ABB RAPID module: Module1.mod

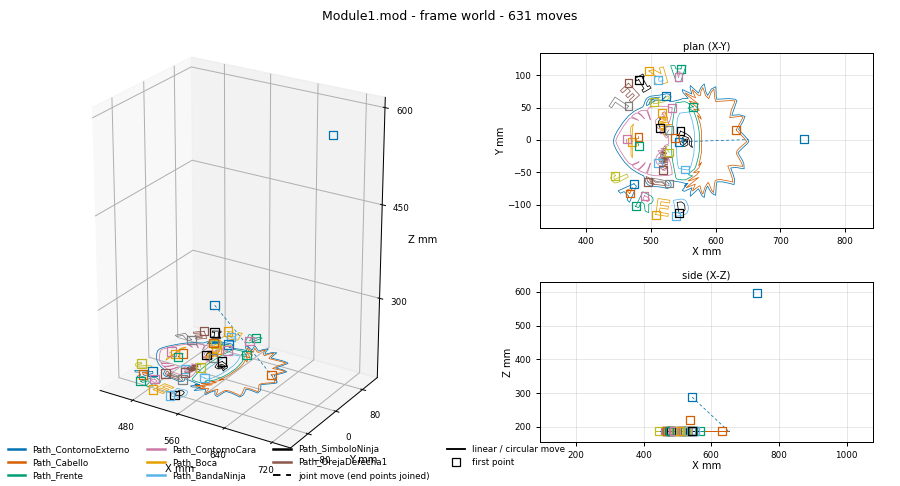
[picture p0: tool path of Module1.mod in frame world, 631 of 636 moves have a stored position in this frame; points joined in program order, loops and branches not executed]
MODULE Module1
    TASK PERS wobjdata Workobject_1:=[FALSE,TRUE,"",[[472.139180242,2.803580658,186.5],[0,0.573617827,0.819123061,0]],[[0,0,0],[1,0,0,0]]];
    TASK PERS wobjdata Cara:=[FALSE,TRUE,"",[[540.229,0.016,186.5],[0,0.707106781,0.707106781,0]],[[0,0,0],[1,0,0,0]]];
    PERS tooldata MyNewTool:=[TRUE,[[8.526,1.82,195.145],[0.965925826,0,0.258819045,0]],[0.14,[0,0,1],[1,0,0,0],0,0,0]];
    CONST robtarget Target_10:=[[-45.629166667,12.05,-2],[0.71519384,0,0,-0.698926156],[0,0,0,0],[9E+09,9E+09,9E+09,9E+09,9E+09,9E+09]];
    CONST robtarget Target_20:=[[-46.396458333,17.381354167,-2],[0.71519384,0,0,-0.698926156],[0,0,0,0],[9E+09,9E+09,9E+09,9E+09,9E+09,9E+09]];
    CONST robtarget Target_30:=[[-42.49468099,20.715104167,-2],[0.71519384,0,0,-0.698926156],[0,0,0,0],[9E+09,9E+09,9E+09,9E+09,9E+09,9E+09]];
    CONST robtarget Target_40:=[[-36.679635417,22.68625,-2],[0.71519384,0,0,-0.698926156],[0,0,0,0],[9E+09,9E+09,9E+09,9E+09,9E+09,9E+09]];
    CONST robtarget Target_50:=[[-21.710833333,26.072916667,-2],[0.71519384,0,0,-0.698926156],[0,0,0,0],[9E+09,9E+09,9E+09,9E+09,9E+09,9E+09]];
    CONST robtarget Target_60:=[[-4.75765625,27.104791667,-2],[0.71519384,0,0,-0.698926156],[0,0,0,0],[9E+09,9E+09,9E+09,9E+09,9E+09,9E+09]];
    CONST robtarget Target_70:=[[12.314583333,26.866666667,-2],[0.71519384,0,0,-0.698926156],[0,0,0,0],[9E+09,9E+09,9E+09,9E+09,9E+09,9E+09]];
    CONST robtarget Target_80:=[[26.688072917,24.458958333,-2],[0.71519384,0,0,-0.698926156],[0,0,0,0],[9E+09,9E+09,9E+09,9E+09,9E+09,9E+09]];
    CONST robtarget Target_90:=[[39.6725,20.46375,-2],[0.71519384,0,0,-0.698926156],[0,0,0,0],[9E+09,9E+09,9E+09,9E+09,9E+09,9E+09]];
    CONST robtarget Target_100:=[[43.257604167,18.849791667,-2],[0.71519384,0,0,-0.698926156],[0,0,0,0],[9E+09,9E+09,9E+09,9E+09,9E+09,9E+09]];
    CONST robtarget Target_110:=[[41.365833333,4.27125,-2],[0.71519384,0,0,-0.698926156],[0,0,0,0],[9E+09,9E+09,9E+09,9E+09,9E+09,9E+09]];
    CONST robtarget Target_120:=[[32.581666667,0.567083333,-2],[0.71519384,0,0,-0.698926156],[0,0,0,0],[9E+09,9E+09,9E+09,9E+09,9E+09,9E+09]];
    CONST robtarget Target_130:=[[22.252167969,-0.135716146,-2],[0.71519384,0,0,-0.698926156],[0,0,0,0],[9E+09,9E+09,9E+09,9E+09,9E+09,9E+09]];
    CONST robtarget Target_140:=[[-12.892766927,-0.549127604,-2],[0.71519384,0,0,-0.698926156],[0,0,0,0],[9E+09,9E+09,9E+09,9E+09,9E+09,9E+09]];
    CONST robtarget Target_150:=[[-26.05,-0.120833333,-2],[0.71519384,0,0,-0.698926156],[0,0,0,0],[9E+09,9E+09,9E+09,9E+09,9E+09,9E+09]];
    CONST robtarget Target_160:=[[-37.334479167,1.129322917,-2],[0.71519384,0,0,-0.698926156],[0,0,0,0],[9E+09,9E+09,9E+09,9E+09,9E+09,9E+09]];
    CONST robtarget Target_170:=[[-43.618333333,2.577916667,-2],[0.71519384,0,0,-0.698926156],[0,0,0,0],[9E+09,9E+09,9E+09,9E+09,9E+09,9E+09]];
    CONST robtarget Target_180:=[[-45.629166667,12.05,-2],[0.71519384,0,0,-0.698926156],[0,0,0,0],[9E+09,9E+09,9E+09,9E+09,9E+09,9E+09]];
    CONST robtarget Target_190:=[[0.514166667,109.68125,-2],[0.71519384,0,0,-0.698926156],[0,0,0,0],[9E+09,9E+09,9E+09,9E+09,9E+09,9E+09]];
    CONST robtarget Target_200:=[[16.547916667,95.129166667,-2],[0.71519384,0,0,-0.698926156],[0,0,0,0],[9E+09,9E+09,9E+09,9E+09,9E+09,9E+09]];
    CONST robtarget Target_210:=[[29.843229167,102.623489583,-2],[0.71519384,0,0,-0.698926156],[0,0,0,0],[9E+09,9E+09,9E+09,9E+09,9E+09,9E+09]];
    CONST robtarget Target_220:=[[36.33875,105.024583333,-2],[0.71519384,0,0,-0.698926156],[0,0,0,0],[9E+09,9E+09,9E+09,9E+09,9E+09,9E+09]];
    CONST robtarget Target_230:=[[38.865520833,96.729895833,-2],[0.71519384,0,0,-0.698926156],[0,0,0,0],[9E+09,9E+09,9E+09,9E+09,9E+09,9E+09]];
    CONST robtarget Target_240:=[[38.06515625,84.664895833,-2],[0.71519384,0,0,-0.698926156],[0,0,0,0],[9E+09,9E+09,9E+09,9E+09,9E+09,9E+09]];
    CONST robtarget Target_250:=[[60.680416667,92.642083333,-2],[0.71519384,0,0,-0.698926156],[0,0,0,0],[9E+09,9E+09,9E+09,9E+09,9E+09,9E+09]];
    CONST robtarget Target_260:=[[62.955833333,89.308333333,-2],[0.71519384,0,0,-0.698926156],[0,0,0,0],[9E+09,9E+09,9E+09,9E+09,9E+09,9E+09]];
    CONST robtarget Target_270:=[[63.82234375,79.750260417,-2],[0.71519384,0,0,-0.698926156],[0,0,0,0],[9E+09,9E+09,9E+09,9E+09,9E+09,9E+09]];
    CONST robtarget Target_280:=[[62.797083333,61.632916667,-2],[0.71519384,0,0,-0.698926156],[0,0,0,0],[9E+09,9E+09,9E+09,9E+09,9E+09,9E+09]];
    CONST robtarget Target_290:=[[67.427291667,60.640729167,-2],[0.71519384,0,0,-0.698926156],[0,0,0,0],[9E+09,9E+09,9E+09,9E+09,9E+09,9E+09]];
    CONST robtarget Target_300:=[[82.15796875,60.058645833,-2],[0.71519384,0,0,-0.698926156],[0,0,0,0],[9E+09,9E+09,9E+09,9E+09,9E+09,9E+09]];
    CONST robtarget Target_310:=[[78.797760417,53.338229167,-2],[0.71519384,0,0,-0.698926156],[0,0,0,0],[9E+09,9E+09,9E+09,9E+09,9E+09,9E+09]];
    CONST robtarget Target_320:=[[68.670833333,47.398333333,-2],[0.71519384,0,0,-0.698926156],[0,0,0,0],[9E+09,9E+09,9E+09,9E+09,9E+09,9E+09]];
    CONST robtarget Target_330:=[[74.352760417,44.5540625,-2],[0.71519384,0,0,-0.698926156],[0,0,0,0],[9E+09,9E+09,9E+09,9E+09,9E+09,9E+09]];
    CONST robtarget Target_340:=[[86.345,42.318333333,-2],[0.71519384,0,0,-0.698926156],[0,0,0,0],[9E+09,9E+09,9E+09,9E+09,9E+09,9E+09]];
    CONST robtarget Target_350:=[[84.1621875,39.53359375,-2],[0.71519384,0,0,-0.698926156],[0,0,0,0],[9E+09,9E+09,9E+09,9E+09,9E+09,9E+09]];
    CONST robtarget Target_360:=[[79.51875,36.232916667,-2],[0.71519384,0,0,-0.698926156],[0,0,0,0],[9E+09,9E+09,9E+09,9E+09,9E+09,9E+09]];
    CONST robtarget Target_370:=[[72.375,33.3225,-2],[0.71519384,0,0,-0.698926156],[0,0,0,0],[9E+09,9E+09,9E+09,9E+09,9E+09,9E+09]];
    CONST robtarget Target_380:=[[84.016666667,20.569583333,-2],[0.71519384,0,0,-0.698926156],[0,0,0,0],[9E+09,9E+09,9E+09,9E+09,9E+09,9E+09]];
    CONST robtarget Target_390:=[[80.821822917,20.331458333,-2],[0.71519384,0,0,-0.698926156],[0,0,0,0],[9E+09,9E+09,9E+09,9E+09,9E+09,9E+09]];
    CONST robtarget Target_400:=[[70.94625,22.950833333,-2],[0.71519384,0,0,-0.698926156],[0,0,0,0],[9E+09,9E+09,9E+09,9E+09,9E+09,9E+09]];
    CONST robtarget Target_410:=[[77.746041667,8.385520833,-2],[0.71519384,0,0,-0.698926156],[0,0,0,0],[9E+09,9E+09,9E+09,9E+09,9E+09,9E+09]];
    CONST robtarget Target_420:=[[73.598697917,9.146197917,-2],[0.71519384,0,0,-0.698926156],[0,0,0,0],[9E+09,9E+09,9E+09,9E+09,9E+09,9E+09]];
    CONST robtarget Target_430:=[[64.172916667,17.394583333,-2],[0.71519384,0,0,-0.698926156],[0,0,0,0],[9E+09,9E+09,9E+09,9E+09,9E+09,9E+09]];
    CONST robtarget Target_440:=[[63.736354167,8.65671875,-2],[0.71519384,0,0,-0.698926156],[0,0,0,0],[9E+09,9E+09,9E+09,9E+09,9E+09,9E+09]];
    CONST robtarget Target_450:=[[62.000852865,4.113326823,-2],[0.71519384,0,0,-0.698926156],[0,0,0,0],[9E+09,9E+09,9E+09,9E+09,9E+09,9E+09]];
    CONST robtarget Target_460:=[[59.28391276,-7.539915365,-2],[0.71519384,0,0,-0.698926156],[0,0,0,0],[9E+09,9E+09,9E+09,9E+09,9E+09,9E+09]];
    CONST robtarget Target_470:=[[58.987083333,-11.074583333,-2],[0.71519384,0,0,-0.698926156],[0,0,0,0],[9E+09,9E+09,9E+09,9E+09,9E+09,9E+09]];
    CONST robtarget Target_480:=[[66.7790625,-9.156354167,-2],[0.71519384,0,0,-0.698926156],[0,0,0,0],[9E+09,9E+09,9E+09,9E+09,9E+09,9E+09]];
    CONST robtarget Target_490:=[[70.522916667,-12.027083333,-2],[0.715023643,0.015246994,0.015601871,-0.69875983],[0,0,0,0],[9E+09,9E+09,9E+09,9E+09,9E+09,9E+09]];
    CONST robtarget Target_500:=[[71.26375,-15.744479167,-2],[0.714513134,0.030486731,0.031196317,-0.698260933],[0,0,0,0],[9E+09,9E+09,9E+09,9E+09,9E+09,9E+09]];
    CONST robtarget Target_510:=[[69.391822917,-25.586979167,-2],[0.713662555,0.045711958,0.046775915,-0.697429701],[0,0,0,0],[9E+09,9E+09,9E+09,9E+09,9E+09,9E+09]];
    CONST robtarget Target_520:=[[67.380989583,-41.475208333,-2],[0.712472311,0.060915428,0.06233325,-0.696266531],[0,0,0,0],[9E+09,9E+09,9E+09,9E+09,9E+09,9E+09]];
    CONST robtarget Target_530:=[[64.490416667,-46.158333333,-2],[0.712472311,0.060915428,0.06233325,-0.696266531],[0,0,0,0],[9E+09,9E+09,9E+09,9E+09,9E+09,9E+09]];
    CONST robtarget Target_540:=[[61.67921875,-48.387447917,-2],[0.712472311,0.060915428,0.06233325,-0.696266531],[0,0,0,0],[9E+09,9E+09,9E+09,9E+09,9E+09,9E+09]];
    CONST robtarget Target_550:=[[54.350260417,-51.03328125,-2],[0.712472311,0.060915428,0.06233325,-0.696266531],[0,0,0,0],[9E+09,9E+09,9E+09,9E+09,9E+09,9E+09]];
    CONST robtarget Target_560:=[[51.214947917,-52.409114583,-2],[0.710942969,0.076089906,0.077860918,-0.694771976],[0,0,0,0],[9E+09,9E+09,9E+09,9E+09,9E+09,9E+09]];
    CONST robtarget Target_570:=[[44.472207031,-65.71186849,-2],[0.710942969,0.076089906,0.077860918,-0.694771976],[0,0,0,0],[9E+09,9E+09,9E+09,9E+09,9E+09,9E+09]];
    CONST robtarget Target_580:=[[37.364010417,-74.52828125,-2],[0.710942969,0.076089906,0.077860918,-0.694771976],[0,0,0,0],[9E+09,9E+09,9E+09,9E+09,9E+09,9E+09]];
    CONST robtarget Target_590:=[[27.586829427,-82.957740885,-2],[0.706870064,0.106323014,0.108797708,-0.690791712],[0,0,0,0],[9E+09,9E+09,9E+09,9E+09,9E+09,9E+09]];
    CONST robtarget Target_600:=[[14.43125,-91.719583333,-2],[0.709075257,0.09122817,0.093351528,-0.692946746],[0,0,0,0],[9E+09,9E+09,9E+09,9E+09,9E+09,9E+09]];
    CONST robtarget Target_610:=[[5.091458333,-96.535,-2],[0.709075257,0.09122817,0.093351528,-0.692946746],[0,0,0,0],[9E+09,9E+09,9E+09,9E+09,9E+09,9E+09]];
    CONST robtarget Target_620:=[[-1.867083333,-98.016666667,-2],[0.709075257,0.09122817,0.093351528,-0.692946746],[0,0,0,0],[9E+09,9E+09,9E+09,9E+09,9E+09,9E+09]];
    CONST robtarget Target_630:=[[-7.6746875,-97.037708333,-2],[0.709075257,0.09122817,0.093351528,-0.692946746],[0,0,0,0],[9E+09,9E+09,9E+09,9E+09,9E+09,9E+09]];
    CONST robtarget Target_640:=[[-16.101666667,-93.095416667,-2],[0.709075257,0.09122817,0.093351528,-0.692946746],[0,0,0,0],[9E+09,9E+09,9E+09,9E+09,9E+09,9E+09]];
    CONST robtarget Target_650:=[[-24.727083333,-87.6846875,-2],[0.709075257,0.09122817,0.093351528,-0.692946746],[0,0,0,0],[9E+09,9E+09,9E+09,9E+09,9E+09,9E+09]];
    CONST robtarget Target_660:=[[-35.09875,-80.130833333,-2],[0.710942969,0.076089907,0.077860918,-0.694771976],[0,0,0,0],[9E+09,9E+09,9E+09,9E+09,9E+09,9E+09]];
    CONST robtarget Target_670:=[[-44.36578125,-70.652135417,-2],[0.712472311,0.060915428,0.06233325,-0.696266531],[0,0,0,0],[9E+09,9E+09,9E+09,9E+09,9E+09,9E+09]];
    CONST robtarget Target_680:=[[-50.97375,-60.34,-2],[0.712472311,0.060915428,0.06233325,-0.696266531],[0,0,0,0],[9E+09,9E+09,9E+09,9E+09,9E+09,9E+09]];
    CONST robtarget Target_690:=[[-55.41875,-51.29125,-2],[0.712989136,0.054837114,0.056113461,-0.6967716],[0,0,0,0],[9E+09,9E+09,9E+09,9E+09,9E+09,9E+09]];
    CONST robtarget Target_700:=[[-66.055,-47.434947917,-2],[0.712989136,0.054837114,0.05611346,-0.6967716],[0,0,0,0],[9E+09,9E+09,9E+09,9E+09,9E+09,9E+09]];
    CONST robtarget Target_710:=[[-69.124166667,-44.570833333,-2],[0.713662554,0.045711958,0.046775915,-0.697429702],[0,0,0,0],[9E+09,9E+09,9E+09,9E+09,9E+09,9E+09]];
    CONST robtarget Target_720:=[[-71.03578125,-40.092760417,-2],[0.714513134,0.030486731,0.031196317,-0.698260933],[0,0,0,0],[9E+09,9E+09,9E+09,9E+09,9E+09,9E+09]];
    CONST robtarget Target_730:=[[-72.735729167,-24.707239583,-2],[0.71519384,0,0,-0.698926156],[0,0,0,0],[9E+09,9E+09,9E+09,9E+09,9E+09,9E+09]];
    CONST robtarget Target_740:=[[-74.733333333,-14.9375,-2],[0.71519384,0,0,-0.698926156],[0,0,0,0],[9E+09,9E+09,9E+09,9E+09,9E+09,9E+09]];
    CONST robtarget Target_750:=[[-73.57578125,-11.312708333,-2],[0.71519384,0,0,-0.698926156],[0,0,0,0],[9E+09,9E+09,9E+09,9E+09,9E+09,9E+09]];
    CONST robtarget Target_760:=[[-71.029166667,-8.957916667,-2],[0.71519384,0,0,-0.698926156],[0,0,0,0],[9E+09,9E+09,9E+09,9E+09,9E+09,9E+09]];
    CONST robtarget Target_770:=[[-67.4440625,-9.1034375,-2],[0.71519384,0,0,-0.698926156],[0,0,0,0],[9E+09,9E+09,9E+09,9E+09,9E+09,9E+09]];
    CONST robtarget Target_780:=[[-63.03875,-11.7625,-2],[0.71519384,0,0,-0.698926156],[0,0,0,0],[9E+09,9E+09,9E+09,9E+09,9E+09,9E+09]];
    CONST robtarget Target_790:=[[-62.873385417,-8.045104167,-2],[0.71519384,0,0,-0.698926156],[0,0,0,0],[9E+09,9E+09,9E+09,9E+09,9E+09,9E+09]];
    CONST robtarget Target_800:=[[-65.347239583,7.22796875,-2],[0.71519384,0,0,-0.698926156],[0,0,0,0],[9E+09,9E+09,9E+09,9E+09,9E+09,9E+09]];
    CONST robtarget Target_810:=[[-66.795833333,11.838333333,-2],[0.71519384,0,0,-0.698926156],[0,0,0,0],[9E+09,9E+09,9E+09,9E+09,9E+09,9E+09]];
    CONST robtarget Target_820:=[[-67.272083333,15.225,-2],[0.71519384,0,0,-0.698926156],[0,0,0,0],[9E+09,9E+09,9E+09,9E+09,9E+09,9E+09]];
    CONST robtarget Target_830:=[[-71.29375,11.785416667,-2],[0.71519384,0,0,-0.698926156],[0,0,0,0],[9E+09,9E+09,9E+09,9E+09,9E+09,9E+09]];
    CONST robtarget Target_840:=[[-66.4915625,17.024166667,-2],[0.71519384,0,0,-0.698926156],[0,0,0,0],[9E+09,9E+09,9E+09,9E+09,9E+09,9E+09]];
    CONST robtarget Target_850:=[[-77.769427083,8.286302083,-2],[0.71519384,0,0,-0.698926156],[0,0,0,0],[9E+09,9E+09,9E+09,9E+09,9E+09,9E+09]];
    CONST robtarget Target_860:=[[-79.264322917,11.408385417,-2],[0.71519384,0,0,-0.698926156],[0,0,0,0],[9E+09,9E+09,9E+09,9E+09,9E+09,9E+09]];
    CONST robtarget Target_870:=[[-73.780833333,23.1625,-2],[0.71519384,0,0,-0.698926156],[0,0,0,0],[9E+09,9E+09,9E+09,9E+09,9E+09,9E+09]];
    CONST robtarget Target_880:=[[-81.923385417,20.609270833,-2],[0.71519384,0,0,-0.698926156],[0,0,0,0],[9E+09,9E+09,9E+09,9E+09,9E+09,9E+09]];
    CONST robtarget Target_890:=[[-86.904166667,20.6225,-2],[0.71519384,0,0,-0.698926156],[0,0,0,0],[9E+09,9E+09,9E+09,9E+09,9E+09,9E+09]];
    CONST robtarget Target_900:=[[-75.2625,33.269583333,-2],[0.71519384,0,0,-0.698926156],[0,0,0,0],[9E+09,9E+09,9E+09,9E+09,9E+09,9E+09]];
    CONST robtarget Target_910:=[[-86.203020833,38.7596875,-2],[0.71519384,0,0,-0.698926156],[0,0,0,0],[9E+09,9E+09,9E+09,9E+09,9E+09,9E+09]];
    CONST robtarget Target_920:=[[-88.809166667,42.159583333,-2],[0.71519384,0,0,-0.698926156],[0,0,0,0],[9E+09,9E+09,9E+09,9E+09,9E+09,9E+09]];
    CONST robtarget Target_930:=[[-80.170520833,43.555260417,-2],[0.71519384,0,0,-0.698926156],[0,0,0,0],[9E+09,9E+09,9E+09,9E+09,9E+09,9E+09]];
    CONST robtarget Target_940:=[[-73.9925,45.599166667,-2],[0.71519384,0,0,-0.698926156],[0,0,0,0],[9E+09,9E+09,9E+09,9E+09,9E+09,9E+09]];
    CONST robtarget Target_950:=[[-71.23421875,47.2528125,-2],[0.71519384,0,0,-0.698926156],[0,0,0,0],[9E+09,9E+09,9E+09,9E+09,9E+09,9E+09]];
    CONST robtarget Target_960:=[[-76.479583333,50.077239583,-2],[0.71519384,0,0,-0.698926156],[0,0,0,0],[9E+09,9E+09,9E+09,9E+09,9E+09,9E+09]];
    CONST robtarget Target_970:=[[-81.506666667,53.272083333,-2],[0.71519384,0,0,-0.698926156],[0,0,0,0],[9E+09,9E+09,9E+09,9E+09,9E+09,9E+09]];
    CONST robtarget Target_980:=[[-84.026822917,56.665364583,-2],[0.71519384,0,0,-0.698926156],[0,0,0,0],[9E+09,9E+09,9E+09,9E+09,9E+09,9E+09]];
    CONST robtarget Target_990:=[[-85.316666667,59.622083333,-2],[0.71519384,0,0,-0.698926156],[0,0,0,0],[9E+09,9E+09,9E+09,9E+09,9E+09,9E+09]];
    CONST robtarget Target_1000:=[[-78.860833333,60.15125,-2],[0.71519384,0,0,-0.698926156],[0,0,0,0],[9E+09,9E+09,9E+09,9E+09,9E+09,9E+09]];
    CONST robtarget Target_1010:=[[-69.501197917,60.706875,-2],[0.71519384,0,0,-0.698926156],[0,0,0,0],[9E+09,9E+09,9E+09,9E+09,9E+09,9E+09]];
    CONST robtarget Target_1020:=[[-64.62625,61.8975,-2],[0.71519384,0,0,-0.698926156],[0,0,0,0],[9E+09,9E+09,9E+09,9E+09,9E+09,9E+09]];
    CONST robtarget Target_1030:=[[-64.619635417,70.126041667,-2],[0.71519384,0,0,-0.698926156],[0,0,0,0],[9E+09,9E+09,9E+09,9E+09,9E+09,9E+09]];
    CONST robtarget Target_1040:=[[-67.272083333,82.323333333,-2],[0.71519384,0,0,-0.698926156],[0,0,0,0],[9E+09,9E+09,9E+09,9E+09,9E+09,9E+09]];
    CONST robtarget Target_1050:=[[-68.9125,87.985416667,-2],[0.71519384,0,0,-0.698926156],[0,0,0,0],[9E+09,9E+09,9E+09,9E+09,9E+09,9E+09]];
    CONST robtarget Target_1060:=[[-62.297916667,89.149583333,-2],[0.71519384,0,0,-0.698926156],[0,0,0,0],[9E+09,9E+09,9E+09,9E+09,9E+09,9E+09]];
    CONST robtarget Target_1070:=[[-54.677916667,87.2975,-2],[0.71519384,0,0,-0.698926156],[0,0,0,0],[9E+09,9E+09,9E+09,9E+09,9E+09,9E+09]];
    CONST robtarget Target_1080:=[[-43.280989583,82.95171875,-2],[0.71519384,0,0,-0.698926156],[0,0,0,0],[9E+09,9E+09,9E+09,9E+09,9E+09,9E+09]];
    CONST robtarget Target_1090:=[[-42.275572917,90.479114583,-2],[0.71519384,0,0,-0.698926156],[0,0,0,0],[9E+09,9E+09,9E+09,9E+09,9E+09,9E+09]];
    CONST robtarget Target_1100:=[[-44.570833333,103.754583333,-2],[0.71519384,0,0,-0.698926156],[0,0,0,0],[9E+09,9E+09,9E+09,9E+09,9E+09,9E+09]];
    CONST robtarget Target_1110:=[[-36.633333333,103.278333333,-2],[0.71519384,0,0,-0.698926156],[0,0,0,0],[9E+09,9E+09,9E+09,9E+09,9E+09,9E+09]];
    CONST robtarget Target_1120:=[[-31.381354167,101.055833333,-2],[0.71519384,0,0,-0.698926156],[0,0,0,0],[9E+09,9E+09,9E+09,9E+09,9E+09,9E+09]];
    CONST robtarget Target_1130:=[[-19.752916667,94.070833333,-2],[0.71519384,0,0,-0.698926156],[0,0,0,0],[9E+09,9E+09,9E+09,9E+09,9E+09,9E+09]];
    CONST robtarget Target_1140:=[[-13.918854167,99.69984375,-2],[0.71519384,0,0,-0.698926156],[0,0,0,0],[9E+09,9E+09,9E+09,9E+09,9E+09,9E+09]];
    CONST robtarget Target_1150:=[[-6.259166667,107.987916667,-2],[0.71519384,0,0,-0.698926156],[0,0,0,0],[9E+09,9E+09,9E+09,9E+09,9E+09,9E+09]];
    CONST robtarget Target_1160:=[[-2.93203125,110.858645833,-2],[0.71519384,0,0,-0.698926156],[0,0,0,0],[9E+09,9E+09,9E+09,9E+09,9E+09,9E+09]];
    CONST robtarget Target_1170:=[[0.514166667,109.68125,-2],[0.71519384,0,0,-0.698926156],[0,0,0,0],[9E+09,9E+09,9E+09,9E+09,9E+09,9E+09]];
    CONST robtarget Target_1350:=[[15.489583333,91.425,-2],[0.71519384,0,0,-0.698926156],[0,0,0,0],[9E+09,9E+09,9E+09,9E+09,9E+09,9E+09]];
    CONST robtarget Target_1360:=[[34.94389974,101.979394531,-2],[0.71519384,0,0,-0.698926156],[0,0,0,0],[9E+09,9E+09,9E+09,9E+09,9E+09,9E+09]];
    CONST robtarget Target_1370:=[[36.669479167,98.674583333,-2],[0.71519384,0,0,-0.698926156],[0,0,0,0],[9E+09,9E+09,9E+09,9E+09,9E+09,9E+09]];
    CONST robtarget Target_1380:=[[34.321302083,81.436979167,-2],[0.71519384,0,0,-0.698926156],[0,0,0,0],[9E+09,9E+09,9E+09,9E+09,9E+09,9E+09]];
    CONST robtarget Target_1390:=[[46.763333333,84.016666667,-2],[0.71519384,0,0,-0.698926156],[0,0,0,0],[9E+09,9E+09,9E+09,9E+09,9E+09,9E+09]];
    CONST robtarget Target_1400:=[[56.129583333,88.177239583,-2],[0.71519384,0,0,-0.698926156],[0,0,0,0],[9E+09,9E+09,9E+09,9E+09,9E+09,9E+09]];
    CONST robtarget Target_1410:=[[60.257083333,89.52,-2],[0.71519384,0,0,-0.698926156],[0,0,0,0],[9E+09,9E+09,9E+09,9E+09,9E+09,9E+09]];
    CONST robtarget Target_1420:=[[60.706875,81.291458333,-2],[0.71519384,0,0,-0.698926156],[0,0,0,0],[9E+09,9E+09,9E+09,9E+09,9E+09,9E+09]];
    CONST robtarget Target_1430:=[[59.304583333,59.886666667,-2],[0.71519384,0,0,-0.698926156],[0,0,0,0],[9E+09,9E+09,9E+09,9E+09,9E+09,9E+09]];
    CONST robtarget Target_1440:=[[63.8025,58.56375,-2],[0.71519384,0,0,-0.698926156],[0,0,0,0],[9E+09,9E+09,9E+09,9E+09,9E+09,9E+09]];
    CONST robtarget Target_1450:=[[78.725,57.029166667,-2],[0.71519384,0,0,-0.698926156],[0,0,0,0],[9E+09,9E+09,9E+09,9E+09,9E+09,9E+09]];
    CONST robtarget Target_1460:=[[73.48625,52.84875,-2],[0.71519384,0,0,-0.698926156],[0,0,0,0],[9E+09,9E+09,9E+09,9E+09,9E+09,9E+09]];
    CONST robtarget Target_1470:=[[63.709895833,49.151197917,-2],[0.71519384,0,0,-0.698926156],[0,0,0,0],[9E+09,9E+09,9E+09,9E+09,9E+09,9E+09]];
    CONST robtarget Target_1480:=[[68.50546875,44.21671875,-2],[0.71519384,0,0,-0.698926156],[0,0,0,0],[9E+09,9E+09,9E+09,9E+09,9E+09,9E+09]];
    CONST robtarget Target_1490:=[[80.861510417,40.042916667,-2],[0.71519384,0,0,-0.698926156],[0,0,0,0],[9E+09,9E+09,9E+09,9E+09,9E+09,9E+09]];
    CONST robtarget Target_1500:=[[75.655833333,37.238333333,-2],[0.71519384,0,0,-0.698926156],[0,0,0,0],[9E+09,9E+09,9E+09,9E+09,9E+09,9E+09]];
    CONST robtarget Target_1510:=[[68.466608073,36.107239583,-2],[0.71519384,0,0,-0.698926156],[0,0,0,0],[9E+09,9E+09,9E+09,9E+09,9E+09,9E+09]];
    CONST robtarget Target_1520:=[[69.142949219,32.819791667,-2],[0.71519384,0,0,-0.698926156],[0,0,0,0],[9E+09,9E+09,9E+09,9E+09,9E+09,9E+09]];
    CONST robtarget Target_1530:=[[77.507916667,23.850416667,-2],[0.71519384,0,0,-0.698926156],[0,0,0,0],[9E+09,9E+09,9E+09,9E+09,9E+09,9E+09]];
    CONST robtarget Target_1540:=[[74.504895833,24.544947917,-2],[0.71519384,0,0,-0.698926156],[0,0,0,0],[9E+09,9E+09,9E+09,9E+09,9E+09,9E+09]];
    CONST robtarget Target_1550:=[[65.0725,28.771666667,-2],[0.71519384,0,0,-0.698926156],[0,0,0,0],[9E+09,9E+09,9E+09,9E+09,9E+09,9E+09]];
    CONST robtarget Target_1560:=[[67.03703125,24.128229167,-2],[0.71519384,0,0,-0.698926156],[0,0,0,0],[9E+09,9E+09,9E+09,9E+09,9E+09,9E+09]];
    CONST robtarget Target_1570:=[[72.6925,12.685,-2],[0.71519384,0,0,-0.698926156],[0,0,0,0],[9E+09,9E+09,9E+09,9E+09,9E+09,9E+09]];
    CONST robtarget Target_1580:=[[69.028020833,15.992291667,-2],[0.71519384,0,0,-0.698926156],[0,0,0,0],[9E+09,9E+09,9E+09,9E+09,9E+09,9E+09]];
    CONST robtarget Target_1590:=[[55.124166667,33.587083333,-2],[0.71519384,0,0,-0.698926156],[0,0,0,0],[9E+09,9E+09,9E+09,9E+09,9E+09,9E+09]];
    CONST robtarget Target_1600:=[[60.376145833,19.008541667,-2],[0.71519384,0,0,-0.698926156],[0,0,0,0],[9E+09,9E+09,9E+09,9E+09,9E+09,9E+09]];
    CONST robtarget Target_1610:=[[57.267291667,21.660989583,-2],[0.71519384,0,0,-0.698926156],[0,0,0,0],[9E+09,9E+09,9E+09,9E+09,9E+09,9E+09]];
    CONST robtarget Target_1620:=[[53.272083333,27.554583333,-2],[0.71519384,0,0,-0.698926156],[0,0,0,0],[9E+09,9E+09,9E+09,9E+09,9E+09,9E+09]];
    CONST robtarget Target_1630:=[[48.787395833,32.297239583,-2],[0.71519384,0,0,-0.698926156],[0,0,0,0],[9E+09,9E+09,9E+09,9E+09,9E+09,9E+09]];
    CONST robtarget Target_1640:=[[45.652083333,34.698333333,-2],[0.71519384,0,0,-0.698926156],[0,0,0,0],[9E+09,9E+09,9E+09,9E+09,9E+09,9E+09]];
    CONST robtarget Target_1650:=[[47.656302083,25.771126302,-2],[0.71519384,0,0,-0.698926156],[0,0,0,0],[9E+09,9E+09,9E+09,9E+09,9E+09,9E+09]];
    CONST robtarget Target_1660:=[[41.471666667,32.581666667,-2],[0.71519384,0,0,-0.698926156],[0,0,0,0],[9E+09,9E+09,9E+09,9E+09,9E+09,9E+09]];
    CONST robtarget Target_1670:=[[36.18,36.193229167,-2],[0.71519384,0,0,-0.698926156],[0,0,0,0],[9E+09,9E+09,9E+09,9E+09,9E+09,9E+09]];
    CONST robtarget Target_1680:=[[31.957725423,37.723368327,-2],[0.71519384,0,0,-0.698926156],[0,0,0,0],[9E+09,9E+09,9E+09,9E+09,9E+09,9E+09]];
    CONST robtarget Target_1690:=[[38.137916667,31.787916667,-2],[0.71519384,0,0,-0.698926156],[0,0,0,0],[9E+09,9E+09,9E+09,9E+09,9E+09,9E+09]];
    CONST robtarget Target_1700:=[[24.262174479,36.184960938,-2],[0.71519384,0,0,-0.698926156],[0,0,0,0],[9E+09,9E+09,9E+09,9E+09,9E+09,9E+09]];
    CONST robtarget Target_1710:=[[11.282708333,38.2040625,-2],[0.71519384,0,0,-0.698926156],[0,0,0,0],[9E+09,9E+09,9E+09,9E+09,9E+09,9E+09]];
    CONST robtarget Target_1720:=[[-18.377083333,37.92625,-2],[0.71519384,0,0,-0.698926156],[0,0,0,0],[9E+09,9E+09,9E+09,9E+09,9E+09,9E+09]];
    CONST robtarget Target_1730:=[[-27.955,36.265989583,-2],[0.71519384,0,0,-0.698926156],[0,0,0,0],[9E+09,9E+09,9E+09,9E+09,9E+09,9E+09]];
    CONST robtarget Target_1740:=[[-39.328052572,33.621809896,-2],[0.71519384,0,0,-0.698926156],[0,0,0,0],[9E+09,9E+09,9E+09,9E+09,9E+09,9E+09]];
    CONST robtarget Target_1750:=[[-34.252083333,38.085,-2],[0.71519384,0,0,-0.698926156],[0,0,0,0],[9E+09,9E+09,9E+09,9E+09,9E+09,9E+09]];
    CONST robtarget Target_1760:=[[-42.851041667,34.01703125,-2],[0.71519384,0,0,-0.698926156],[0,0,0,0],[9E+09,9E+09,9E+09,9E+09,9E+09,9E+09]];
    CONST robtarget Target_1770:=[[-50.644054362,25.739603678,-2],[0.71519384,0,0,-0.698926156],[0,0,0,0],[9E+09,9E+09,9E+09,9E+09,9E+09,9E+09]];
    CONST robtarget Target_1780:=[[-48.539583333,34.698333333,-2],[0.71519384,0,0,-0.698926156],[0,0,0,0],[9E+09,9E+09,9E+09,9E+09,9E+09,9E+09]];
    CONST robtarget Target_1790:=[[-53.6725,30.729583333,-2],[0.71519384,0,0,-0.698926156],[0,0,0,0],[9E+09,9E+09,9E+09,9E+09,9E+09,9E+09]];
    CONST robtarget Target_1800:=[[-61.329707031,20.051165365,-2],[0.71519384,0,0,-0.698926156],[0,0,0,0],[9E+09,9E+09,9E+09,9E+09,9E+09,9E+09]];
    CONST robtarget Target_1810:=[[-62.9990625,17.354895833,-2],[0.71519384,0,0,-0.698926156],[0,0,0,0],[9E+09,9E+09,9E+09,9E+09,9E+09,9E+09]];
    CONST robtarget Target_1820:=[[-62.78078125,20.64234375,-2],[0.71519384,0,0,-0.698926156],[0,0,0,0],[9E+09,9E+09,9E+09,9E+09,9E+09,9E+09]];
    CONST robtarget Target_1830:=[[-57.890020345,33.671419271,-2],[0.71519384,0,0,-0.698926156],[0,0,0,0],[9E+09,9E+09,9E+09,9E+09,9E+09,9E+09]];
    CONST robtarget Target_1840:=[[-71.141614583,17.163072917,-2],[0.71519384,0,0,-0.698926156],[0,0,0,0],[9E+09,9E+09,9E+09,9E+09,9E+09,9E+09]];
    CONST robtarget Target_1850:=[[-73.87922526,14.268365885,-2],[0.71519384,0,0,-0.698926156],[0,0,0,0],[9E+09,9E+09,9E+09,9E+09,9E+09,9E+09]];
    CONST robtarget Target_1860:=[[-70.215572917,23.030208333,-2],[0.71519384,0,0,-0.698926156],[0,0,0,0],[9E+09,9E+09,9E+09,9E+09,9E+09,9E+09]];
    CONST robtarget Target_1870:=[[-68.184895833,28.407864583,-2],[0.71519384,0,0,-0.698926156],[0,0,0,0],[9E+09,9E+09,9E+09,9E+09,9E+09,9E+09]];
    CONST robtarget Target_1880:=[[-78.65578125,24.088541667,-2],[0.71519384,0,0,-0.698926156],[0,0,0,0],[9E+09,9E+09,9E+09,9E+09,9E+09,9E+09]];
    CONST robtarget Target_1890:=[[-72.080885417,32.7271875,-2],[0.71519384,0,0,-0.698926156],[0,0,0,0],[9E+09,9E+09,9E+09,9E+09,9E+09,9E+09]];
    CONST robtarget Target_1900:=[[-70.65875,35.650833333,-2],[0.71519384,0,0,-0.698926156],[0,0,0,0],[9E+09,9E+09,9E+09,9E+09,9E+09,9E+09]];
    CONST robtarget Target_1910:=[[-80.018385417,37.979166667,-2],[0.71519384,0,0,-0.698926156],[0,0,0,0],[9E+09,9E+09,9E+09,9E+09,9E+09,9E+09]];
    CONST robtarget Target_1920:=[[-83.570416667,39.884166667,-2],[0.71519384,0,0,-0.698926156],[0,0,0,0],[9E+09,9E+09,9E+09,9E+09,9E+09,9E+09]];
    CONST robtarget Target_1930:=[[-72.041197917,43.74046875,-2],[0.71519384,0,0,-0.698926156],[0,0,0,0],[9E+09,9E+09,9E+09,9E+09,9E+09,9E+09]];
    CONST robtarget Target_1940:=[[-65.26125,48.192083333,-2],[0.71519384,0,0,-0.698926156],[0,0,0,0],[9E+09,9E+09,9E+09,9E+09,9E+09,9E+09]];
    CONST robtarget Target_1950:=[[-68.965416667,50.15,-2],[0.71519384,0,0,-0.698926156],[0,0,0,0],[9E+09,9E+09,9E+09,9E+09,9E+09,9E+09]];
    CONST robtarget Target_1960:=[[-77.564375,53.589583333,-2],[0.71519384,0,0,-0.698926156],[0,0,0,0],[9E+09,9E+09,9E+09,9E+09,9E+09,9E+09]];
    CONST robtarget Target_1970:=[[-81.244150391,56.486150716,-2],[0.71519384,0,0,-0.698926156],[0,0,0,0],[9E+09,9E+09,9E+09,9E+09,9E+09,9E+09]];
    CONST robtarget Target_1980:=[[-67.42421875,58.02796875,-2],[0.71519384,0,0,-0.698926156],[0,0,0,0],[9E+09,9E+09,9E+09,9E+09,9E+09,9E+09]];
    CONST robtarget Target_1990:=[[-63.144583333,59.145833333,-2],[0.71519384,0,0,-0.698926156],[0,0,0,0],[9E+09,9E+09,9E+09,9E+09,9E+09,9E+09]];
    CONST robtarget Target_2000:=[[-61.466959635,61.796627604,-2],[0.71519384,0,0,-0.698926156],[0,0,0,0],[9E+09,9E+09,9E+09,9E+09,9E+09,9E+09]];
    CONST robtarget Target_2010:=[[-60.95515625,66.7790625,-2],[0.71519384,0,0,-0.698926156],[0,0,0,0],[9E+09,9E+09,9E+09,9E+09,9E+09,9E+09]];
    CONST robtarget Target_2020:=[[-63.409166667,80.206666667,-2],[0.71519384,0,0,-0.698926156],[0,0,0,0],[9E+09,9E+09,9E+09,9E+09,9E+09,9E+09]];
    CONST robtarget Target_2030:=[[-65.049583333,86.50375,-2],[0.71519384,0,0,-0.698926156],[0,0,0,0],[9E+09,9E+09,9E+09,9E+09,9E+09,9E+09]];
    CONST robtarget Target_2040:=[[-58.408541667,85.240364583,-2],[0.71519384,0,0,-0.698926156],[0,0,0,0],[9E+09,9E+09,9E+09,9E+09,9E+09,9E+09]];
    CONST robtarget Target_2050:=[[-47.9575,81.635416667,-2],[0.71519384,0,0,-0.698926156],[0,0,0,0],[9E+09,9E+09,9E+09,9E+09,9E+09,9E+09]];
    CONST robtarget Target_2060:=[[-40.258125,78.42734375,-2],[0.71519384,0,0,-0.698926156],[0,0,0,0],[9E+09,9E+09,9E+09,9E+09,9E+09,9E+09]];
    CONST robtarget Target_2070:=[[-38.80953125,85.743072917,-2],[0.71519384,0,0,-0.698926156],[0,0,0,0],[9E+09,9E+09,9E+09,9E+09,9E+09,9E+09]];
    CONST robtarget Target_2080:=[[-40.81375,101.796666667,-2],[0.71519384,0,0,-0.698926156],[0,0,0,0],[9E+09,9E+09,9E+09,9E+09,9E+09,9E+09]];
    CONST robtarget Target_2090:=[[-35.389791667,99.68,-2],[0.71519384,0,0,-0.698926156],[0,0,0,0],[9E+09,9E+09,9E+09,9E+09,9E+09,9E+09]];
    CONST robtarget Target_2100:=[[-21.492552083,91.92109375,-2],[0.71519384,0,0,-0.698926156],[0,0,0,0],[9E+09,9E+09,9E+09,9E+09,9E+09,9E+09]];
    CONST robtarget Target_2110:=[[-16.706074219,92.589166667,-2],[0.71519384,0,0,-0.698926156],[0,0,0,0],[9E+09,9E+09,9E+09,9E+09,9E+09,9E+09]];
    CONST robtarget Target_2120:=[[-12.787760417,96.121354167,-2],[0.71519384,0,0,-0.698926156],[0,0,0,0],[9E+09,9E+09,9E+09,9E+09,9E+09,9E+09]];
    CONST robtarget Target_2130:=[[-2.555,107.829166667,-2],[0.71519384,0,0,-0.698926156],[0,0,0,0],[9E+09,9E+09,9E+09,9E+09,9E+09,9E+09]];
    CONST robtarget Target_2140:=[[2.604375,103.90671875,-2],[0.71519384,0,0,-0.698926156],[0,0,0,0],[9E+09,9E+09,9E+09,9E+09,9E+09,9E+09]];
    CONST robtarget Target_2150:=[[15.489583333,91.425,-2],[0.71519384,0,0,-0.698926156],[0,0,0,0],[9E+09,9E+09,9E+09,9E+09,9E+09,9E+09]];
    CONST robtarget Target_2160:=[[13.690416667,5.488333333,-2],[0.71519384,0,0,-0.698926156],[0,0,0,0],[9E+09,9E+09,9E+09,9E+09,9E+09,9E+09]];
    CONST robtarget Target_2170:=[[9.404166667,14.854583333,-2],[0.71519384,0,0,-0.698926156],[0,0,0,0],[9E+09,9E+09,9E+09,9E+09,9E+09,9E+09]];
    CONST robtarget Target_2180:=[[5.547864583,19.855208333,-2],[0.71519384,0,0,-0.698926156],[0,0,0,0],[9E+09,9E+09,9E+09,9E+09,9E+09,9E+09]];
    CONST robtarget Target_2190:=[[1.89,22.315833333,-2],[0.71519384,0,0,-0.698926156],[0,0,0,0],[9E+09,9E+09,9E+09,9E+09,9E+09,9E+09]];
    CONST robtarget Target_2200:=[[-1.3246875,23.116197917,-2],[0.71519384,0,0,-0.698926156],[0,0,0,0],[9E+09,9E+09,9E+09,9E+09,9E+09,9E+09]];
    CONST robtarget Target_2210:=[[-7.25796875,22.216614583,-2],[0.71519384,0,0,-0.698926156],[0,0,0,0],[9E+09,9E+09,9E+09,9E+09,9E+09,9E+09]];
    CONST robtarget Target_2220:=[[-11.539257813,24.157994792,-2],[0.71519384,0,0,-0.698926156],[0,0,0,0],[9E+09,9E+09,9E+09,9E+09,9E+09,9E+09]];
    CONST robtarget Target_2230:=[[-9.8575,21.151666667,-2],[0.71519384,0,0,-0.698926156],[0,0,0,0],[9E+09,9E+09,9E+09,9E+09,9E+09,9E+09]];
    CONST robtarget Target_2240:=[[-6.973541667,19.01515625,-2],[0.71519384,0,0,-0.698926156],[0,0,0,0],[9E+09,9E+09,9E+09,9E+09,9E+09,9E+09]];
    CONST robtarget Target_2250:=[[-2.502083333,19.458333333,-2],[0.71519384,0,0,-0.698926156],[0,0,0,0],[9E+09,9E+09,9E+09,9E+09,9E+09,9E+09]];
    CONST robtarget Target_2260:=[[3.325364583,17.837760417,-2],[0.71519384,0,0,-0.698926156],[0,0,0,0],[9E+09,9E+09,9E+09,9E+09,9E+09,9E+09]];
    CONST robtarget Target_2270:=[[5.54125,12.05,-2],[0.71519384,0,0,-0.698926156],[0,0,0,0],[9E+09,9E+09,9E+09,9E+09,9E+09,9E+09]];
    CONST robtarget Target_2280:=[[4.01328125,8.703020833,-2],[0.71519384,0,0,-0.698926156],[0,0,0,0],[9E+09,9E+09,9E+09,9E+09,9E+09,9E+09]];
    CONST robtarget Target_2290:=[[-0.49125,7.816666667,-2],[0.71519384,0,0,-0.698926156],[0,0,0,0],[9E+09,9E+09,9E+09,9E+09,9E+09,9E+09]];
    CONST robtarget Target_2300:=[[-3.593489583,8.068020833,-2],[0.71519384,0,0,-0.698926156],[0,0,0,0],[9E+09,9E+09,9E+09,9E+09,9E+09,9E+09]];
    CONST robtarget Target_2310:=[[-7,12.05,-2],[0.71519384,0,0,-0.698926156],[0,0,0,0],[9E+09,9E+09,9E+09,9E+09,9E+09,9E+09]];
    CONST robtarget Target_2320:=[[-2.71375,15.754166667,-2],[0.71519384,0,0,-0.698926156],[0,0,0,0],[9E+09,9E+09,9E+09,9E+09,9E+09,9E+09]];
    CONST robtarget Target_2330:=[[0.00484375,13.564739583,-2],[0.71519384,0,0,-0.698926156],[0,0,0,0],[9E+09,9E+09,9E+09,9E+09,9E+09,9E+09]];
    CONST robtarget Target_2340:=[[-1.92,11.0975,-2],[0.71519384,0,0,-0.698926156],[0,0,0,0],[9E+09,9E+09,9E+09,9E+09,9E+09,9E+09]];
    CONST robtarget Target_2350:=[[1.083020833,10.766770833,-2],[0.71519384,0,0,-0.698926156],[0,0,0,0],[9E+09,9E+09,9E+09,9E+09,9E+09,9E+09]];
    CONST robtarget Target_2360:=[[1.31453125,16.389166667,-2],[0.71519384,0,0,-0.698926156],[0,0,0,0],[9E+09,9E+09,9E+09,9E+09,9E+09,9E+09]];
    CONST robtarget Target_2370:=[[-7.271197917,16.885260417,-2],[0.71519384,0,0,-0.698926156],[0,0,0,0],[9E+09,9E+09,9E+09,9E+09,9E+09,9E+09]];
    CONST robtarget Target_2380:=[[-10.175,11.997083333,-2],[0.71519384,0,0,-0.698926156],[0,0,0,0],[9E+09,9E+09,9E+09,9E+09,9E+09,9E+09]];
    CONST robtarget Target_2390:=[[-7.033072917,5.772760417,-2],[0.71519384,0,0,-0.698926156],[0,0,0,0],[9E+09,9E+09,9E+09,9E+09,9E+09,9E+09]];
    CONST robtarget Target_2400:=[[2.101666667,3.16,-2],[0.71519384,0,0,-0.698926156],[0,0,0,0],[9E+09,9E+09,9E+09,9E+09,9E+09,9E+09]];
    CONST robtarget Target_2410:=[[9.146197917,3.689166667,-2],[0.71519384,0,0,-0.698926156],[0,0,0,0],[9E+09,9E+09,9E+09,9E+09,9E+09,9E+09]];
    CONST robtarget Target_2420:=[[13.690416667,5.488333333,-2],[0.71519384,0,0,-0.698926156],[0,0,0,0],[9E+09,9E+09,9E+09,9E+09,9E+09,9E+09]];
    CONST robtarget Target_2430:=[[51.155416667,25.279166667,-2],[0.71519384,0,0,-0.698926156],[0,0,0,0],[9E+09,9E+09,9E+09,9E+09,9E+09,9E+09]];
    CONST robtarget Target_2440:=[[54.145208333,21.422864583,-2],[0.71519384,0,0,-0.698926156],[0,0,0,0],[9E+09,9E+09,9E+09,9E+09,9E+09,9E+09]];
    CONST robtarget Target_2450:=[[57.92875,15.5425,-2],[0.71519384,0,0,-0.698926156],[0,0,0,0],[9E+09,9E+09,9E+09,9E+09,9E+09,9E+09]];
    CONST robtarget Target_2460:=[[59.145833333,11.467916667,-2],[0.71519384,0,0,-0.698926156],[0,0,0,0],[9E+09,9E+09,9E+09,9E+09,9E+09,9E+09]];
    CONST robtarget Target_2470:=[[57.346666667,-1.6025,-2],[0.71519384,0,0,-0.698926156],[0,0,0,0],[9E+09,9E+09,9E+09,9E+09,9E+09,9E+09]];
    CONST robtarget Target_2480:=[[38.772916667,-5.147916667,-2],[0.71519384,0,0,-0.698926156],[0,0,0,0],[9E+09,9E+09,9E+09,9E+09,9E+09,9E+09]];
    CONST robtarget Target_2490:=[[20.615885417,-7.383645833,-2],[0.71519384,0,0,-0.698926156],[0,0,0,0],[9E+09,9E+09,9E+09,9E+09,9E+09,9E+09]];
    CONST robtarget Target_2500:=[[0.514166667,-8.42875,-2],[0.71519384,0,0,-0.698926156],[0,0,0,0],[9E+09,9E+09,9E+09,9E+09,9E+09,9E+09]];
    CONST robtarget Target_2510:=[[-21.82328125,-7.93265625,-2],[0.71519384,0,0,-0.698926156],[0,0,0,0],[9E+09,9E+09,9E+09,9E+09,9E+09,9E+09]];
    CONST robtarget Target_2520:=[[-32.443821615,-6.605605469,-2],[0.71519384,0,0,-0.698926156],[0,0,0,0],[9E+09,9E+09,9E+09,9E+09,9E+09,9E+09]];
    CONST robtarget Target_2530:=[[-57.74046875,-1.814166667,-2],[0.71519384,0,0,-0.698926156],[0,0,0,0],[9E+09,9E+09,9E+09,9E+09,9E+09,9E+09]];
    CONST robtarget Target_2540:=[[-60.287083333,-0.120833333,-2],[0.71519384,0,0,-0.698926156],[0,0,0,0],[9E+09,9E+09,9E+09,9E+09,9E+09,9E+09]];
    CONST robtarget Target_2550:=[[-61.457864583,6.685572917,-2],[0.71519384,0,0,-0.698926156],[0,0,0,0],[9E+09,9E+09,9E+09,9E+09,9E+09,9E+09]];
    CONST robtarget Target_2560:=[[-61.557083333,13.531666667,-2],[0.71519384,0,0,-0.698926156],[0,0,0,0],[9E+09,9E+09,9E+09,9E+09,9E+09,9E+09]];
    CONST robtarget Target_2570:=[[-55.410481771,24.128229167,-2],[0.71519384,0,0,-0.698926156],[0,0,0,0],[9E+09,9E+09,9E+09,9E+09,9E+09,9E+09]];
    CONST robtarget Target_2580:=[[-53.659270833,17.844375,-2],[0.71519384,0,0,-0.698926156],[0,0,0,0],[9E+09,9E+09,9E+09,9E+09,9E+09,9E+09]];
    CONST robtarget Target_2590:=[[-50.391666667,20.093333333,-2],[0.71519384,0,0,-0.698926156],[0,0,0,0],[9E+09,9E+09,9E+09,9E+09,9E+09,9E+09]];
    CONST robtarget Target_2600:=[[-45.166145833,26.91296875,-2],[0.71519384,0,0,-0.698926156],[0,0,0,0],[9E+09,9E+09,9E+09,9E+09,9E+09,9E+09]];
    CONST robtarget Target_2610:=[[-41.000611979,29.03046224,-2],[0.71519384,0,0,-0.698926156],[0,0,0,0],[9E+09,9E+09,9E+09,9E+09,9E+09,9E+09]];
    CONST robtarget Target_2620:=[[-26.241822917,33.1240625,-2],[0.71519384,0,0,-0.698926156],[0,0,0,0],[9E+09,9E+09,9E+09,9E+09,9E+09,9E+09]];
    CONST robtarget Target_2630:=[[-17.107083333,34.539583333,-2],[0.71519384,0,0,-0.698926156],[0,0,0,0],[9E+09,9E+09,9E+09,9E+09,9E+09,9E+09]];
    CONST robtarget Target_2640:=[[3.646998698,35.246516927,-2],[0.71519384,0,0,-0.698926156],[0,0,0,0],[9E+09,9E+09,9E+09,9E+09,9E+09,9E+09]];
    CONST robtarget Target_2650:=[[15.489583333,33.9575,-2],[0.71519384,0,0,-0.698926156],[0,0,0,0],[9E+09,9E+09,9E+09,9E+09,9E+09,9E+09]];
    CONST robtarget Target_2660:=[[28.546770833,31.364583333,-2],[0.71519384,0,0,-0.698926156],[0,0,0,0],[9E+09,9E+09,9E+09,9E+09,9E+09,9E+09]];
    CONST robtarget Target_2670:=[[39.460833333,27.819166667,-2],[0.71519384,0,0,-0.698926156],[0,0,0,0],[9E+09,9E+09,9E+09,9E+09,9E+09,9E+09]];
    CONST robtarget Target_2680:=[[44.382083333,25.649583333,-2],[0.71519384,0,0,-0.698926156],[0,0,0,0],[9E+09,9E+09,9E+09,9E+09,9E+09,9E+09]];
    CONST robtarget Target_2690:=[[49.303333333,17.077083333,-2],[0.71519384,0,0,-0.698926156],[0,0,0,0],[9E+09,9E+09,9E+09,9E+09,9E+09,9E+09]];
    CONST robtarget Target_2700:=[[51.155416667,25.279166667,-2],[0.71519384,0,0,-0.698926156],[0,0,0,0],[9E+09,9E+09,9E+09,9E+09,9E+09,9E+09]];
    CONST robtarget Target_2710:=[[49.567916667,-7.47625,-2],[0.715023643,0.015246994,0.015601871,-0.69875983],[0,0,0,0],[9E+09,9E+09,9E+09,9E+09,9E+09,9E+09]];
    CONST robtarget Target_2720:=[[51.036354167,-13.118489583,-2],[0.714513134,0.030486731,0.031196317,-0.698260933],[0,0,0,0],[9E+09,9E+09,9E+09,9E+09,9E+09,9E+09]];
    CONST robtarget Target_2730:=[[52.107916667,-23.404166667,-2],[0.713662555,0.045711958,0.046775915,-0.697429701],[0,0,0,0],[9E+09,9E+09,9E+09,9E+09,9E+09,9E+09]];
    CONST robtarget Target_2740:=[[51.115729167,-37.810729167,-2],[0.712472311,0.060915428,0.06233325,-0.696266531],[0,0,0,0],[9E+09,9E+09,9E+09,9E+09,9E+09,9E+09]];
    CONST robtarget Target_2750:=[[49.815963542,-43.376901042,-2],[0.712472311,0.060915428,0.06233325,-0.696266531],[0,0,0,0],[9E+09,9E+09,9E+09,9E+09,9E+09,9E+09]];
    CONST robtarget Target_2760:=[[45.86375,-45.311666667,-2],[0.712472311,0.060915428,0.06233325,-0.696266531],[0,0,0,0],[9E+09,9E+09,9E+09,9E+09,9E+09,9E+09]];
    CONST robtarget Target_2770:=[[36.259375,-41.898541667,-2],[0.712472311,0.060915428,0.06233325,-0.696266531],[0,0,0,0],[9E+09,9E+09,9E+09,9E+09,9E+09,9E+09]];
    CONST robtarget Target_2780:=[[30.99644043,-41.005572917,-2],[0.712472311,0.060915428,0.06233325,-0.696266531],[0,0,0,0],[9E+09,9E+09,9E+09,9E+09,9E+09,9E+09]];
    CONST robtarget Target_2790:=[[38.3628125,-43.823385417,-2],[0.712472311,0.060915428,0.06233325,-0.696266531],[0,0,0,0],[9E+09,9E+09,9E+09,9E+09,9E+09,9E+09]];
    CONST robtarget Target_2800:=[[45.440416667,-46.793333333,-2],[0.712472311,0.060915428,0.06233325,-0.696266531],[0,0,0,0],[9E+09,9E+09,9E+09,9E+09,9E+09,9E+09]];
    CONST robtarget Target_2810:=[[45.374270833,-54.995416667,-2],[0.712472311,0.060915428,0.06233325,-0.696266531],[0,0,0,0],[9E+09,9E+09,9E+09,9E+09,9E+09,9E+09]];
    CONST robtarget Target_2820:=[[42.68875,-59.916666667,-2],[0.712472311,0.060915428,0.06233325,-0.696266531],[0,0,0,0],[9E+09,9E+09,9E+09,9E+09,9E+09,9E+09]];
    CONST robtarget Target_2830:=[[38.376041667,-54.492708333,-2],[0.712472311,0.060915428,0.06233325,-0.696266531],[0,0,0,0],[9E+09,9E+09,9E+09,9E+09,9E+09,9E+09]];
    CONST robtarget Target_2840:=[[33.057916667,-50.18,-2],[0.712472311,0.060915428,0.06233325,-0.696266531],[0,0,0,0],[9E+09,9E+09,9E+09,9E+09,9E+09,9E+09]];
    CONST robtarget Target_2850:=[[37.82703125,-55.365833333,-2],[0.712472311,0.060915428,0.06233325,-0.696266531],[0,0,0,0],[9E+09,9E+09,9E+09,9E+09,9E+09,9E+09]];
    CONST robtarget Target_2860:=[[41.365833333,-60.0225,-2],[0.712472311,0.060915428,0.06233325,-0.696266531],[0,0,0,0],[9E+09,9E+09,9E+09,9E+09,9E+09,9E+09]];
    CONST robtarget Target_2870:=[[41.312916667,-63.35625,-2],[0.712472311,0.060915428,0.06233325,-0.696266531],[0,0,0,0],[9E+09,9E+09,9E+09,9E+09,9E+09,9E+09]];
    CONST robtarget Target_2880:=[[38.428958333,-67.397760417,-2],[0.712472311,0.060915428,0.06233325,-0.696266531],[0,0,0,0],[9E+09,9E+09,9E+09,9E+09,9E+09,9E+09]];
    CONST robtarget Target_2890:=[[35.8625,-69.970833333,-2],[0.712472311,0.060915428,0.06233325,-0.696266531],[0,0,0,0],[9E+09,9E+09,9E+09,9E+09,9E+09,9E+09]];
    CONST robtarget Target_2900:=[[33.315885417,-63.878802083,-2],[0.712472311,0.060915428,0.06233325,-0.696266531],[0,0,0,0],[9E+09,9E+09,9E+09,9E+09,9E+09,9E+09]];
    CONST robtarget Target_2910:=[[30.118147786,-58.911663411,-2],[0.712472311,0.060915428,0.06233325,-0.696266531],[0,0,0,0],[9E+09,9E+09,9E+09,9E+09,9E+09,9E+09]];
    CONST robtarget Target_2920:=[[34.069947917,-69.613645833,-2],[0.712472311,0.060915428,0.06233325,-0.696266531],[0,0,0,0],[9E+09,9E+09,9E+09,9E+09,9E+09,9E+09]];
    CONST robtarget Target_2930:=[[33.428333333,-73.04,-2],[0.712472311,0.060915428,0.06233325,-0.696266531],[0,0,0,0],[9E+09,9E+09,9E+09,9E+09,9E+09,9E+09]];
    CONST robtarget Target_2940:=[[21.27734375,-82.452552083,-2],[0.710942969,0.076089906,0.077860918,-0.694771976],[0,0,0,0],[9E+09,9E+09,9E+09,9E+09,9E+09,9E+09]];
    CONST robtarget Target_2950:=[[6.387916667,-91.190416667,-2],[0.709075257,0.09122817,0.093351528,-0.692946746],[0,0,0,0],[9E+09,9E+09,9E+09,9E+09,9E+09,9E+09]];
    CONST robtarget Target_2960:=[[1.334375,-93.604739583,-2],[0.709075257,0.09122817,0.093351528,-0.692946746],[0,0,0,0],[9E+09,9E+09,9E+09,9E+09,9E+09,9E+09]];
    CONST robtarget Target_2970:=[[-1.655416667,-94.3125,-2],[0.709075257,0.09122817,0.093351528,-0.692946746],[0,0,0,0],[9E+09,9E+09,9E+09,9E+09,9E+09,9E+09]];
    CONST robtarget Target_2980:=[[-7.838398438,-92.16358724,-2],[0.709075257,0.09122817,0.093351528,-0.692946746],[0,0,0,0],[9E+09,9E+09,9E+09,9E+09,9E+09,9E+09]];
    CONST robtarget Target_2990:=[[-17.583333333,-86.924010417,-2],[0.709075257,0.09122817,0.093351528,-0.692946746],[0,0,0,0],[9E+09,9E+09,9E+09,9E+09,9E+09,9E+09]];
    CONST robtarget Target_3000:=[[-27.804518229,-80.404511719,-2],[0.710942969,0.076089906,0.077860918,-0.694771976],[0,0,0,0],[9E+09,9E+09,9E+09,9E+09,9E+09,9E+09]];
    CONST robtarget Target_3010:=[[-35.41625,-74.415833333,-2],[0.712472311,0.060915428,0.06233325,-0.696266531],[0,0,0,0],[9E+09,9E+09,9E+09,9E+09,9E+09,9E+09]];
    CONST robtarget Target_3020:=[[-38.207604167,-69.838541667,-2],[0.712472311,0.060915428,0.06233325,-0.696266531],[0,0,0,0],[9E+09,9E+09,9E+09,9E+09,9E+09,9E+09]];
    CONST robtarget Target_3030:=[[-33.67,-58.27625,-2],[0.712472311,0.060915428,0.06233325,-0.696266531],[0,0,0,0],[9E+09,9E+09,9E+09,9E+09,9E+09,9E+09]];
    CONST robtarget Target_3040:=[[-36.30921875,-62.258229167,-2],[0.712472311,0.060915428,0.06233325,-0.696266531],[0,0,0,0],[9E+09,9E+09,9E+09,9E+09,9E+09,9E+09]];
    CONST robtarget Target_3050:=[[-39.358541667,-68.85296875,-2],[0.712472311,0.060915428,0.06233325,-0.696266531],[0,0,0,0],[9E+09,9E+09,9E+09,9E+09,9E+09,9E+09]];
    CONST robtarget Target_3060:=[[-43.09578125,-65.644895833,-2],[0.712472311,0.060915428,0.06233325,-0.696266531],[0,0,0,0],[9E+09,9E+09,9E+09,9E+09,9E+09,9E+09]];
    CONST robtarget Target_3070:=[[-45.629166667,-60.975,-2],[0.712472311,0.060915428,0.06233325,-0.696266531],[0,0,0,0],[9E+09,9E+09,9E+09,9E+09,9E+09,9E+09]];
    CONST robtarget Target_3080:=[[-43.2346875,-57.098854167,-2],[0.712472311,0.060915428,0.06233325,-0.696266531],[0,0,0,0],[9E+09,9E+09,9E+09,9E+09,9E+09,9E+09]];
    CONST robtarget Target_3090:=[[-35.050380859,-48.920645345,-2],[0.712472311,0.060915428,0.06233325,-0.696266531],[0,0,0,0],[9E+09,9E+09,9E+09,9E+09,9E+09,9E+09]];
    CONST robtarget Target_3100:=[[-37.95625,-50.603333333,-2],[0.712472311,0.060915428,0.06233325,-0.696266531],[0,0,0,0],[9E+09,9E+09,9E+09,9E+09,9E+09,9E+09]];
    CONST robtarget Target_3110:=[[-42.096979167,-54.155364583,-2],[0.712472311,0.060915428,0.06233325,-0.696266531],[0,0,0,0],[9E+09,9E+09,9E+09,9E+09,9E+09,9E+09]];
    CONST robtarget Target_3120:=[[-46.52875,-59.652083333,-2],[0.712472311,0.060915428,0.06233325,-0.696266531],[0,0,0,0],[9E+09,9E+09,9E+09,9E+09,9E+09,9E+09]];
    CONST robtarget Target_3130:=[[-50.424739583,-51.000208333,-2],[0.712472311,0.060915428,0.06233325,-0.696266531],[0,0,0,0],[9E+09,9E+09,9E+09,9E+09,9E+09,9E+09]];
    CONST robtarget Target_3140:=[[-51.1325,-47.64,-2],[0.712472311,0.060915428,0.06233325,-0.696266531],[0,0,0,0],[9E+09,9E+09,9E+09,9E+09,9E+09,9E+09]];
    CONST robtarget Target_3150:=[[-47.289427083,-45.5365625,-2],[0.712472311,0.060915428,0.06233325,-0.696266531],[0,0,0,0],[9E+09,9E+09,9E+09,9E+09,9E+09,9E+09]];
    CONST robtarget Target_3160:=[[-35.786666667,-41.025416667,-2],[0.712472311,0.060915428,0.06233325,-0.696266531],[0,0,0,0],[9E+09,9E+09,9E+09,9E+09,9E+09,9E+09]];
    CONST robtarget Target_3170:=[[-41.27015625,-42.037447917,-2],[0.715023643,0.015246994,0.015601871,-0.69875983],[0,0,0,0],[9E+09,9E+09,9E+09,9E+09,9E+09,9E+09]];
    CONST robtarget Target_3180:=[[-52.296666667,-46.0525,-2],[0.714513134,0.030486731,0.031196317,-0.698260933],[0,0,0,0],[9E+09,9E+09,9E+09,9E+09,9E+09,9E+09]];
    CONST robtarget Target_3190:=[[-53.937083333,-40.549166667,-2],[0.715023643,0.015246994,0.015601871,-0.69875983],[0,0,0,0],[9E+09,9E+09,9E+09,9E+09,9E+09,9E+09]];
    CONST robtarget Target_3200:=[[-55.127708333,-34.5828125,-2],[0.71519384,0,0,-0.698926156],[0,0,0,0],[9E+09,9E+09,9E+09,9E+09,9E+09,9E+09]];
    CONST robtarget Target_3210:=[[-55.365833333,-25.520833333,-2],[0.71519384,0,0,-0.698926156],[0,0,0,0],[9E+09,9E+09,9E+09,9E+09,9E+09,9E+09]];
    CONST robtarget Target_3220:=[[-54.7440625,-13.35,-2],[0.71519384,0,0,-0.698926156],[0,0,0,0],[9E+09,9E+09,9E+09,9E+09,9E+09,9E+09]];
    CONST robtarget Target_3230:=[[-53.090416667,-7.370416667,-2],[0.71519384,0,0,-0.698926156],[0,0,0,0],[9E+09,9E+09,9E+09,9E+09,9E+09,9E+09]];
    CONST robtarget Target_3240:=[[-46.581666667,-7.740833333,-2],[0.71519384,0,0,-0.698926156],[0,0,0,0],[9E+09,9E+09,9E+09,9E+09,9E+09,9E+09]];
    CONST robtarget Target_3250:=[[-37.627174479,-9.503619792,-2],[0.71519384,0,0,-0.698926156],[0,0,0,0],[9E+09,9E+09,9E+09,9E+09,9E+09,9E+09]];
    CONST robtarget Target_3260:=[[-30.944791667,-11.524375,-2],[0.71519384,0,0,-0.698926156],[0,0,0,0],[9E+09,9E+09,9E+09,9E+09,9E+09,9E+09]];
    CONST robtarget Target_3270:=[[-28.112096354,-13.187942708,-2],[0.71519384,0,0,-0.698926156],[0,0,0,0],[9E+09,9E+09,9E+09,9E+09,9E+09,9E+09]];
    CONST robtarget Target_3280:=[[-38.578020833,-14.811822917,-2],[0.71519384,0,0,-0.698926156],[0,0,0,0],[9E+09,9E+09,9E+09,9E+09,9E+09,9E+09]];
    CONST robtarget Target_3290:=[[-45.25875,-16.577916667,-2],[0.71519384,0,0,-0.698926156],[0,0,0,0],[9E+09,9E+09,9E+09,9E+09,9E+09,9E+09]];
    CONST robtarget Target_3300:=[[-47.236510417,-19.078229167,-2],[0.71519384,0,0,-0.698926156],[0,0,0,0],[9E+09,9E+09,9E+09,9E+09,9E+09,9E+09]];
    CONST robtarget Target_3310:=[[-45.364583333,-23.086666667,-2],[0.71519384,0,0,-0.698926156],[0,0,0,0],[9E+09,9E+09,9E+09,9E+09,9E+09,9E+09]];
    CONST robtarget Target_3320:=[[-43.142083333,-25.520833333,-2],[0.71519384,0,0,-0.698926156],[0,0,0,0],[9E+09,9E+09,9E+09,9E+09,9E+09,9E+09]];
    CONST robtarget Target_3330:=[[-42.890729167,-20.487135417,-2],[0.71519384,0,0,-0.698926156],[0,0,0,0],[9E+09,9E+09,9E+09,9E+09,9E+09,9E+09]];
    CONST robtarget Target_3340:=[[-38.915364583,-19.217135417,-2],[0.71519384,0,0,-0.698926156],[0,0,0,0],[9E+09,9E+09,9E+09,9E+09,9E+09,9E+09]];
    CONST robtarget Target_3350:=[[-40.086145833,-23.820885417,-2],[0.71519384,0,0,-0.698926156],[0,0,0,0],[9E+09,9E+09,9E+09,9E+09,9E+09,9E+09]];
    CONST robtarget Target_3360:=[[-39.54375,-26.949583333,-2],[0.71519384,0,0,-0.698926156],[0,0,0,0],[9E+09,9E+09,9E+09,9E+09,9E+09,9E+09]];
    CONST robtarget Target_3370:=[[-36.61266276,-30.704186198,-2],[0.71519384,0,0,-0.698926156],[0,0,0,0],[9E+09,9E+09,9E+09,9E+09,9E+09,9E+09]];
    CONST robtarget Target_3380:=[[-32.089114583,-32.49921875,-2],[0.71519384,0,0,-0.698926156],[0,0,0,0],[9E+09,9E+09,9E+09,9E+09,9E+09,9E+09]];
    CONST robtarget Target_3390:=[[-27.019863281,-32.180891927,-2],[0.71519384,0,0,-0.698926156],[0,0,0,0],[9E+09,9E+09,9E+09,9E+09,9E+09,9E+09]];
    CONST robtarget Target_3400:=[[-22.451666667,-29.595416667,-2],[0.71519384,0,0,-0.698926156],[0,0,0,0],[9E+09,9E+09,9E+09,9E+09,9E+09,9E+09]];
    CONST robtarget Target_3410:=[[-20.17625,-25.944166667,-2],[0.71519384,0,0,-0.698926156],[0,0,0,0],[9E+09,9E+09,9E+09,9E+09,9E+09,9E+09]];
    CONST robtarget Target_3420:=[[-16.525,-29.44328125,-2],[0.71519384,0,0,-0.698926156],[0,0,0,0],[9E+09,9E+09,9E+09,9E+09,9E+09,9E+09]];
    CONST robtarget Target_3430:=[[-16.472083333,-20.49375,-2],[0.71519384,0,0,-0.698926156],[0,0,0,0],[9E+09,9E+09,9E+09,9E+09,9E+09,9E+09]];
    CONST robtarget Target_3440:=[[-12.959739583,-24.885833333,-2],[0.71519384,0,0,-0.698926156],[0,0,0,0],[9E+09,9E+09,9E+09,9E+09,9E+09,9E+09]];
    CONST robtarget Target_3450:=[[-13.720416667,-21.975416667,-2],[0.71519384,0,0,-0.698926156],[0,0,0,0],[9E+09,9E+09,9E+09,9E+09,9E+09,9E+09]];
    CONST robtarget Target_3460:=[[-8.038489583,-17.642864583,-2],[0.71519384,0,0,-0.698926156],[0,0,0,0],[9E+09,9E+09,9E+09,9E+09,9E+09,9E+09]];
    CONST robtarget Target_3470:=[[-6.365,-12.662083333,-2],[0.71519384,0,0,-0.698926156],[0,0,0,0],[9E+09,9E+09,9E+09,9E+09,9E+09,9E+09]];
    CONST robtarget Target_3480:=[[3.63625,-12.820833333,-2],[0.71519384,0,0,-0.698926156],[0,0,0,0],[9E+09,9E+09,9E+09,9E+09,9E+09,9E+09]];
    CONST robtarget Target_3490:=[[3.265833333,-16.392708333,-2],[0.71519384,0,0,-0.698926156],[0,0,0,0],[9E+09,9E+09,9E+09,9E+09,9E+09,9E+09]];
    CONST robtarget Target_3500:=[[6.010885417,-19.012083333,-2],[0.71519384,0,0,-0.698926156],[0,0,0,0],[9E+09,9E+09,9E+09,9E+09,9E+09,9E+09]];
    CONST robtarget Target_3510:=[[9.66875,-21.161822917,-2],[0.71519384,0,0,-0.698926156],[0,0,0,0],[9E+09,9E+09,9E+09,9E+09,9E+09,9E+09]];
    CONST robtarget Target_3520:=[[9.35125,-25.785416667,-2],[0.71519384,0,0,-0.698926156],[0,0,0,0],[9E+09,9E+09,9E+09,9E+09,9E+09,9E+09]];
    CONST robtarget Target_3530:=[[12.26828125,-21.2478125,-2],[0.71519384,0,0,-0.698926156],[0,0,0,0],[9E+09,9E+09,9E+09,9E+09,9E+09,9E+09]];
    CONST robtarget Target_3540:=[[12.3278125,-26.718072917,-2],[0.71519384,0,0,-0.698926156],[0,0,0,0],[9E+09,9E+09,9E+09,9E+09,9E+09,9E+09]];
    CONST robtarget Target_3550:=[[15.754166667,-23.933333333,-2],[0.71519384,0,0,-0.698926156],[0,0,0,0],[9E+09,9E+09,9E+09,9E+09,9E+09,9E+09]];
    CONST robtarget Target_3560:=[[18.783645833,-29.754166667,-2],[0.71519384,0,0,-0.698926156],[0,0,0,0],[9E+09,9E+09,9E+09,9E+09,9E+09,9E+09]];
    CONST robtarget Target_3570:=[[21.945416667,-32.188333333,-2],[0.71519384,0,0,-0.698926156],[0,0,0,0],[9E+09,9E+09,9E+09,9E+09,9E+09,9E+09]];
    CONST robtarget Target_3580:=[[27.342916667,-32.929166667,-2],[0.71519384,0,0,-0.698926156],[0,0,0,0],[9E+09,9E+09,9E+09,9E+09,9E+09,9E+09]];
    CONST robtarget Target_3590:=[[30.828802083,-32.65796875,-2],[0.71519384,0,0,-0.698926156],[0,0,0,0],[9E+09,9E+09,9E+09,9E+09,9E+09,9E+09]];
    CONST robtarget Target_3600:=[[35.730208333,-26.909895833,-2],[0.71519384,0,0,-0.698926156],[0,0,0,0],[9E+09,9E+09,9E+09,9E+09,9E+09,9E+09]];
    CONST robtarget Target_3610:=[[35.96171875,-20.090260417,-2],[0.71519384,0,0,-0.698926156],[0,0,0,0],[9E+09,9E+09,9E+09,9E+09,9E+09,9E+09]];
    CONST robtarget Target_3620:=[[39.011041667,-20.645885417,-2],[0.71519384,0,0,-0.698926156],[0,0,0,0],[9E+09,9E+09,9E+09,9E+09,9E+09,9E+09]];
    CONST robtarget Target_3630:=[[39.51375,-23.615833333,-2],[0.71519384,0,0,-0.698926156],[0,0,0,0],[9E+09,9E+09,9E+09,9E+09,9E+09,9E+09]];
    CONST robtarget Target_3640:=[[43.766927083,-19.52140625,-2],[0.71519384,0,0,-0.698926156],[0,0,0,0],[9E+09,9E+09,9E+09,9E+09,9E+09,9E+09]];
    CONST robtarget Target_3650:=[[41.789166667,-16.8425,-2],[0.71519384,0,0,-0.698926156],[0,0,0,0],[9E+09,9E+09,9E+09,9E+09,9E+09,9E+09]];
    CONST robtarget Target_3660:=[[35.161354167,-15.016875,-2],[0.71519384,0,0,-0.698926156],[0,0,0,0],[9E+09,9E+09,9E+09,9E+09,9E+09,9E+09]];
    CONST robtarget Target_3670:=[[24.508567708,-13.152389323,-2],[0.71519384,0,0,-0.698926156],[0,0,0,0],[9E+09,9E+09,9E+09,9E+09,9E+09,9E+09]];
    CONST robtarget Target_3680:=[[32.131875,-10.062552083,-2],[0.71519384,0,0,-0.698926156],[0,0,0,0],[9E+09,9E+09,9E+09,9E+09,9E+09,9E+09]];
    CONST robtarget Target_3690:=[[38.772916667,-8.5875,-2],[0.71519384,0,0,-0.698926156],[0,0,0,0],[9E+09,9E+09,9E+09,9E+09,9E+09,9E+09]];
    CONST robtarget Target_3700:=[[46.928697917,-7.49609375,-2],[0.71519384,0,0,-0.698926156],[0,0,0,0],[9E+09,9E+09,9E+09,9E+09,9E+09,9E+09]];
    CONST robtarget Target_3710:=[[49.567916667,-7.47625,-2],[0.71519384,0,0,-0.698926156],[0,0,0,0],[9E+09,9E+09,9E+09,9E+09,9E+09,9E+09]];
    CONST robtarget Target_3720:=[[-2.607916667,-68.9125,-2],[0.712472311,0.060915429,0.06233325,-0.696266531],[0,0,0,0],[9E+09,9E+09,9E+09,9E+09,9E+09,9E+09]];
    CONST robtarget Target_3730:=[[15.5821875,-68.760364583,-2],[0.712472311,0.060915429,0.06233325,-0.696266531],[0,0,0,0],[9E+09,9E+09,9E+09,9E+09,9E+09,9E+09]];
    CONST robtarget Target_3740:=[[21.310416667,-67.854166667,-2],[0.712472311,0.060915429,0.06233325,-0.696266531],[0,0,0,0],[9E+09,9E+09,9E+09,9E+09,9E+09,9E+09]];
    CONST robtarget Target_3750:=[[24.657499186,-66.949829102,-2],[0.712472311,0.060915429,0.06233325,-0.696266531],[0,0,0,0],[9E+09,9E+09,9E+09,9E+09,9E+09,9E+09]];
    CONST robtarget Target_3760:=[[20.14625,-71.022552083,-2],[0.712472311,0.060915429,0.06233325,-0.696266531],[0,0,0,0],[9E+09,9E+09,9E+09,9E+09,9E+09,9E+09]];
    CONST robtarget Target_3770:=[[15.287838542,-71.375605469,-2],[0.712472311,0.060915429,0.06233325,-0.696266531],[0,0,0,0],[9E+09,9E+09,9E+09,9E+09,9E+09,9E+09]];
    CONST robtarget Target_3780:=[[-0.31265625,-70.6190625,-2],[0.712472311,0.060915429,0.06233325,-0.696266531],[0,0,0,0],[9E+09,9E+09,9E+09,9E+09,9E+09,9E+09]];
    CONST robtarget Target_3790:=[[-22.603802083,-70.903489583,-2],[0.712472311,0.060915429,0.06233325,-0.696266531],[0,0,0,0],[9E+09,9E+09,9E+09,9E+09,9E+09,9E+09]];
    CONST robtarget Target_3800:=[[-27.584583333,-68.700833333,-2],[0.712472311,0.060915429,0.06233325,-0.696266531],[0,0,0,0],[9E+09,9E+09,9E+09,9E+09,9E+09,9E+09]];
    CONST robtarget Target_3810:=[[-20.798020833,-68.760364583,-2],[0.712472311,0.060915429,0.06233325,-0.696266531],[0,0,0,0],[9E+09,9E+09,9E+09,9E+09,9E+09,9E+09]];
    CONST robtarget Target_3820:=[[-2.607916667,-68.9125,-2],[0.712472311,0.060915429,0.06233325,-0.696266531],[0,0,0,0],[9E+09,9E+09,9E+09,9E+09,9E+09,9E+09]];
    CONST robtarget Target_3830:=[[-64.573333333,-44.465,-2],[0.713662555,0.045711958,0.046775915,-0.697429701],[0,0,0,0],[9E+09,9E+09,9E+09,9E+09,9E+09,9E+09]];
    CONST robtarget Target_3840:=[[-59.777760417,-46.674270833,-2],[0.713662555,0.045711958,0.046775915,-0.697429701],[0,0,0,0],[9E+09,9E+09,9E+09,9E+09,9E+09,9E+09]];
    CONST robtarget Target_3850:=[[-56.37125,-47.534166667,-2],[0.713662555,0.045711958,0.046775915,-0.697429701],[0,0,0,0],[9E+09,9E+09,9E+09,9E+09,9E+09,9E+09]];
    CONST robtarget Target_3860:=[[-58.223333333,-43.089166667,-2],[0.713662555,0.045711958,0.046775915,-0.697429701],[0,0,0,0],[9E+09,9E+09,9E+09,9E+09,9E+09,9E+09]];
    CONST robtarget Target_3870:=[[-64.24921875,-41.045260417,-2],[0.713662555,0.045711958,0.046775915,-0.697429701],[0,0,0,0],[9E+09,9E+09,9E+09,9E+09,9E+09,9E+09]];
    CONST robtarget Target_3880:=[[-67.219166667,-38.485416667,-2],[0.713662555,0.045711958,0.046775915,-0.697429701],[0,0,0,0],[9E+09,9E+09,9E+09,9E+09,9E+09,9E+09]];
    CONST robtarget Target_3890:=[[-67.854166667,-35.151666667,-2],[0.713662555,0.045711958,0.046775915,-0.697429701],[0,0,0,0],[9E+09,9E+09,9E+09,9E+09,9E+09,9E+09]];
    CONST robtarget Target_3900:=[[-63.819270833,-39.22625,-2],[0.713662555,0.045711958,0.046775915,-0.697429701],[0,0,0,0],[9E+09,9E+09,9E+09,9E+09,9E+09,9E+09]];
    CONST robtarget Target_3910:=[[-59.599166667,-40.866666667,-2],[0.713662555,0.045711958,0.046775915,-0.697429701],[0,0,0,0],[9E+09,9E+09,9E+09,9E+09,9E+09,9E+09]];
    CONST robtarget Target_3920:=[[-65.168645833,-33.220208333,-2],[0.714513134,0.030486731,0.031196317,-0.698260933],[0,0,0,0],[9E+09,9E+09,9E+09,9E+09,9E+09,9E+09]];
    CONST robtarget Target_3930:=[[-65.208333333,-27.531666667,-2],[0.715023643,0.015246994,0.015601871,-0.69875983],[0,0,0,0],[9E+09,9E+09,9E+09,9E+09,9E+09,9E+09]];
    CONST robtarget Target_3940:=[[-64.8246875,-24.257447917,-2],[0.71519384,0,0,-0.698926156],[0,0,0,0],[9E+09,9E+09,9E+09,9E+09,9E+09,9E+09]];
    CONST robtarget Target_3950:=[[-68.039375,-19.5809375,-2],[0.71519384,0,0,-0.698926156],[0,0,0,0],[9E+09,9E+09,9E+09,9E+09,9E+09,9E+09]];
    CONST robtarget Target_3960:=[[-70.489251302,-17.722239583,-2],[0.71519384,0,0,-0.698926156],[0,0,0,0],[9E+09,9E+09,9E+09,9E+09,9E+09,9E+09]];
    CONST robtarget Target_3970:=[[-68.197298177,-36.949179687,-2],[0.715023643,0.015246994,0.015601871,-0.69875983],[0,0,0,0],[9E+09,9E+09,9E+09,9E+09,9E+09,9E+09]];
    CONST robtarget Target_3980:=[[-67.38453125,-40.81375,-2],[0.714513134,0.030486731,0.031196317,-0.698260933],[0,0,0,0],[9E+09,9E+09,9E+09,9E+09,9E+09,9E+09]];
    CONST robtarget Target_3990:=[[-64.573333333,-44.465,-2],[0.714513134,0.030486731,0.031196317,-0.698260933],[0,0,0,0],[9E+09,9E+09,9E+09,9E+09,9E+09,9E+09]];
    CONST robtarget Target_4000:=[[-67.16625,-12.55625,-2],[0.71519384,0,0,-0.698926156],[0,0,0,0],[9E+09,9E+09,9E+09,9E+09,9E+09,9E+09]];
    CONST robtarget Target_4010:=[[-62.965989583,-17.986822917,-2],[0.71519384,0,0,-0.698926156],[0,0,0,0],[9E+09,9E+09,9E+09,9E+09,9E+09,9E+09]];
    CONST robtarget Target_4020:=[[-61.458691406,-23.100722656,-2],[0.71519384,0,0,-0.698926156],[0,0,0,0],[9E+09,9E+09,9E+09,9E+09,9E+09,9E+09]];
    CONST robtarget Target_4030:=[[-58.882311198,-38.484589844,-2],[0.715023643,0.015246994,0.015601871,-0.69875983],[0,0,0,0],[9E+09,9E+09,9E+09,9E+09,9E+09,9E+09]];
    CONST robtarget Target_4040:=[[-62.5625,-34.516666667,-2],[0.71519384,0,0,-0.698926156],[0,0,0,0],[9E+09,9E+09,9E+09,9E+09,9E+09,9E+09]];
    CONST robtarget Target_4050:=[[-63.89203125,-31.7253125,-2],[0.71519384,0,0,-0.698926156],[0,0,0,0],[9E+09,9E+09,9E+09,9E+09,9E+09,9E+09]];
    CONST robtarget Target_4060:=[[-63.462083333,-22.5575,-2],[0.71519384,0,0,-0.698926156],[0,0,0,0],[9E+09,9E+09,9E+09,9E+09,9E+09,9E+09]];
    CONST robtarget Target_4070:=[[-69.494583333,-15.89,-2],[0.71519384,0,0,-0.698926156],[0,0,0,0],[9E+09,9E+09,9E+09,9E+09,9E+09,9E+09]];
    CONST robtarget Target_4080:=[[-70.5,-12.027083333,-2],[0.71519384,0,0,-0.698926156],[0,0,0,0],[9E+09,9E+09,9E+09,9E+09,9E+09,9E+09]];
    CONST robtarget Target_4090:=[[-67.16625,-12.55625,-2],[0.71519384,0,0,-0.698926156],[0,0,0,0],[9E+09,9E+09,9E+09,9E+09,9E+09,9E+09]];
    CONST robtarget Target_4100:=[[58.88125,-35.363333333,-2],[0.71519384,0,0,-0.698926156],[0,0,0,0],[9E+09,9E+09,9E+09,9E+09,9E+09,9E+09]];
    CONST robtarget Target_4110:=[[60.839166667,-32.452916667,-2],[0.71519384,0,0,-0.698926156],[0,0,0,0],[9E+09,9E+09,9E+09,9E+09,9E+09,9E+09]];
    CONST robtarget Target_4120:=[[60.118177083,-25.011510417,-2],[0.71519384,0,0,-0.698926156],[0,0,0,0],[9E+09,9E+09,9E+09,9E+09,9E+09,9E+09]];
    CONST robtarget Target_4130:=[[68.141666667,-13.985,-2],[0.71519384,0,0,-0.698926156],[0,0,0,0],[9E+09,9E+09,9E+09,9E+09,9E+09,9E+09]];
    CONST robtarget Target_4140:=[[65.7075,-11.7625,-2],[0.71519384,0,0,-0.698926156],[0,0,0,0],[9E+09,9E+09,9E+09,9E+09,9E+09,9E+09]];
    CONST robtarget Target_4150:=[[62.320833333,-14.355416667,-2],[0.71519384,0,0,-0.698926156],[0,0,0,0],[9E+09,9E+09,9E+09,9E+09,9E+09,9E+09]];
    CONST robtarget Target_4160:=[[58.874635417,-19.871979167,-2],[0.71519384,0,0,-0.698926156],[0,0,0,0],[9E+09,9E+09,9E+09,9E+09,9E+09,9E+09]];
    CONST robtarget Target_4170:=[[56.5,-31.024166667,-2],[0.71519384,0,0,-0.698926156],[0,0,0,0],[9E+09,9E+09,9E+09,9E+09,9E+09,9E+09]];
    CONST robtarget Target_4180:=[[55.740976563,-36.300950521,-2],[0.71519384,0,0,-0.698926156],[0,0,0,0],[9E+09,9E+09,9E+09,9E+09,9E+09,9E+09]];
    CONST robtarget Target_4190:=[[58.88125,-35.363333333,-2],[0.71519384,0,0,-0.698926156],[0,0,0,0],[9E+09,9E+09,9E+09,9E+09,9E+09,9E+09]];
    CONST robtarget Target_4200:=[[67.665416667,-17.31875,-2],[0.71519384,0,0,-0.698926156],[0,0,0,0],[9E+09,9E+09,9E+09,9E+09,9E+09,9E+09]];
    CONST robtarget Target_4210:=[[64.569791667,-19.845520833,-2],[0.71519384,0,0,-0.698926156],[0,0,0,0],[9E+09,9E+09,9E+09,9E+09,9E+09,9E+09]];
    CONST robtarget Target_4220:=[[61.474166667,-23.562916667,-2],[0.71519384,0,0,-0.698926156],[0,0,0,0],[9E+09,9E+09,9E+09,9E+09,9E+09,9E+09]];
    CONST robtarget Target_4230:=[[61.646145833,-33.498020833,-2],[0.715023643,0.015246994,0.015601871,-0.69875983],[0,0,0,0],[9E+09,9E+09,9E+09,9E+09,9E+09,9E+09]];
    CONST robtarget Target_4240:=[[57.77,-38.485416667,-2],[0.714513134,0.030486731,0.031196317,-0.698260933],[0,0,0,0],[9E+09,9E+09,9E+09,9E+09,9E+09,9E+09]];
    CONST robtarget Target_4250:=[[54.647916667,-41.554583333,-2],[0.714513134,0.030486731,0.031196317,-0.698260933],[0,0,0,0],[9E+09,9E+09,9E+09,9E+09,9E+09,9E+09]];
    CONST robtarget Target_4260:=[[59.727916667,-40.02,-2],[0.714513134,0.030486731,0.031196317,-0.698260933],[0,0,0,0],[9E+09,9E+09,9E+09,9E+09,9E+09,9E+09]];
    CONST robtarget Target_4270:=[[62.420052083,-37.367552083,-2],[0.714513134,0.030486731,0.031196317,-0.698260933],[0,0,0,0],[9E+09,9E+09,9E+09,9E+09,9E+09,9E+09]];
    CONST robtarget Target_4280:=[[64.126614583,-33.187135417,-2],[0.714513134,0.030486731,0.031196317,-0.698260933],[0,0,0,0],[9E+09,9E+09,9E+09,9E+09,9E+09,9E+09]];
    CONST robtarget Target_4290:=[[62.459739583,-40.244895833,-2],[0.714513134,0.030486731,0.031196317,-0.698260933],[0,0,0,0],[9E+09,9E+09,9E+09,9E+09,9E+09,9E+09]];
    CONST robtarget Target_4300:=[[54.409791667,-43.538958333,-2],[0.714513134,0.030486731,0.031196317,-0.698260933],[0,0,0,0],[9E+09,9E+09,9E+09,9E+09,9E+09,9E+09]];
    CONST robtarget Target_4310:=[[52.974427083,-46.760260417,-2],[0.714513134,0.030486731,0.031196317,-0.698260933],[0,0,0,0],[9E+09,9E+09,9E+09,9E+09,9E+09,9E+09]];
    CONST robtarget Target_4320:=[[57.346666667,-46.654427083,-2],[0.714513134,0.030486731,0.031196317,-0.698260933],[0,0,0,0],[9E+09,9E+09,9E+09,9E+09,9E+09,9E+09]];
    CONST robtarget Target_4330:=[[62.479583333,-43.777083333,-2],[0.714513134,0.030486731,0.031196317,-0.698260933],[0,0,0,0],[9E+09,9E+09,9E+09,9E+09,9E+09,9E+09]];
    CONST robtarget Target_4340:=[[64.583020833,-40.264739583,-2],[0.714513134,0.030486731,0.031196317,-0.698260933],[0,0,0,0],[9E+09,9E+09,9E+09,9E+09,9E+09,9E+09]];
    CONST robtarget Target_4350:=[[66.117604167,-26.056614583,-2],[0.714513134,0.030486731,0.031196317,-0.698260933],[0,0,0,0],[9E+09,9E+09,9E+09,9E+09,9E+09,9E+09]];
    CONST robtarget Target_4360:=[[67.665416667,-17.31875,-2],[0.714513134,0.030486731,0.031196317,-0.698260933],[0,0,0,0],[9E+09,9E+09,9E+09,9E+09,9E+09,9E+09]];
    CONST robtarget Target_4490:=[[5.170833333,-59.334583333,-2],[0.712472312,0.060915429,0.06233325,-0.696266531],[0,0,0,0],[9E+09,9E+09,9E+09,9E+09,9E+09,9E+09]];
    CONST robtarget Target_4500:=[[1.995833333,-59.652083333,-2],[0.712472312,0.060915429,0.06233325,-0.696266531],[0,0,0,0],[9E+09,9E+09,9E+09,9E+09,9E+09,9E+09]];
    CONST robtarget Target_4510:=[[2.419166667,-60.445833333,-2],[0.712472312,0.060915429,0.06233325,-0.696266531],[0,0,0,0],[9E+09,9E+09,9E+09,9E+09,9E+09,9E+09]];
    CONST robtarget Target_4520:=[[-8.992,-58.958,-2],[0.712472312,0.060915429,0.06233325,-0.696266531],[0,0,0,0],[9E+09,9E+09,9E+09,9E+09,9E+09,9E+09]];
    CONST robtarget Target_4530:=[[-6.065,-59.24,-2],[0.712472312,0.060915429,0.06233325,-0.696266531],[0,0,0,0],[9E+09,9E+09,9E+09,9E+09,9E+09,9E+09]];
    CONST robtarget Target_4540:=[[-5.738,-60.369,-2],[0.712472312,0.060915429,0.06233325,-0.696266531],[0,0,0,0],[9E+09,9E+09,9E+09,9E+09,9E+09,9E+09]];
    CONST robtarget Target_4550:=[[0.912,-77.305,-2],[0.712472311,0.060915428,0.06233325,-0.696266531],[0,0,0,0],[9E+09,9E+09,9E+09,9E+09,9E+09,9E+09]];
    CONST robtarget Target_4560:=[[-1.715,-77.906,-2],[0.712472311,0.060915428,0.06233325,-0.696266531],[0,0,0,0],[9E+09,9E+09,9E+09,9E+09,9E+09,9E+09]];
    CONST robtarget Target_4570:=[[-4.775,-77.228,-2],[0.712472311,0.060915428,0.06233325,-0.696266531],[0,0,0,0],[9E+09,9E+09,9E+09,9E+09,9E+09,9E+09]];
    CONST robtarget Target_4580:=[[42.242,-22.641,-2],[0.71519384,0,0,-0.698926156],[0,0,0,0],[9E+09,9E+09,9E+09,9E+09,9E+09,9E+09]];
    CONST robtarget Target_4590:=[[40.689,-16.421,-2],[0.71519384,0,0,-0.698926156],[0,0,0,0],[9E+09,9E+09,9E+09,9E+09,9E+09,9E+09]];
    CONST robtarget Target_4600:=[[36.066,-19.892,-2],[0.71519384,0,0,-0.698926156],[0,0,0,0],[9E+09,9E+09,9E+09,9E+09,9E+09,9E+09]];
    CONST robtarget Target_4610:=[[33.871,-14.746,-2],[0.71519384,0,0,-0.698926156],[0,0,0,0],[9E+09,9E+09,9E+09,9E+09,9E+09,9E+09]];
    CONST robtarget Target_4620:=[[32.357,-25.134,-2],[0.71519384,0,0,-0.698926156],[0,0,0,0],[9E+09,9E+09,9E+09,9E+09,9E+09,9E+09]];
    CONST robtarget Target_4630:=[[31.042,-14.218,-2],[0.71519384,0,0,-0.698926156],[0,0,0,0],[9E+09,9E+09,9E+09,9E+09,9E+09,9E+09]];
    CONST robtarget Target_4640:=[[27.408,-29.149,-2],[0.71519384,0,0,-0.698926156],[0,0,0,0],[9E+09,9E+09,9E+09,9E+09,9E+09,9E+09]];
    CONST robtarget Target_4650:=[[27.617,-13.823,-2],[0.71519384,0,0,-0.698926156],[0,0,0,0],[9E+09,9E+09,9E+09,9E+09,9E+09,9E+09]];
    CONST robtarget Target_4660:=[[24.758,-28.49,-2],[0.71519384,0,0,-0.698926156],[0,0,0,0],[9E+09,9E+09,9E+09,9E+09,9E+09,9E+09]];
    CONST robtarget Target_4670:=[[23.867,-7.086,-2],[0.71519384,0,0,-0.698926156],[0,0,0,0],[9E+09,9E+09,9E+09,9E+09,9E+09,9E+09]];
    CONST robtarget Target_4680:=[[21.006,-25.651,-2],[0.71519384,0,0,-0.698926156],[0,0,0,0],[9E+09,9E+09,9E+09,9E+09,9E+09,9E+09]];
    CONST robtarget Target_4690:=[[20.255,-13.477,-2],[0.71519384,0,0,-0.698926156],[0,0,0,0],[9E+09,9E+09,9E+09,9E+09,9E+09,9E+09]];
    CONST robtarget Target_4700:=[[17.047,-26.788,-2],[0.71519384,0,0,-0.698926156],[0,0,0,0],[9E+09,9E+09,9E+09,9E+09,9E+09,9E+09]];
    CONST robtarget Target_4710:=[[16.862,-15.832,-2],[0.71519384,0,0,-0.698926156],[0,0,0,0],[9E+09,9E+09,9E+09,9E+09,9E+09,9E+09]];
    CONST robtarget Target_4720:=[[15.165,-24.693,-2],[0.71519384,0,0,-0.698926156],[0,0,0,0],[9E+09,9E+09,9E+09,9E+09,9E+09,9E+09]];
    CONST robtarget Target_4760:=[[-35.73375,-28.9075,-2],[0.71519384,0,0,-0.698926156],[0,0,0,0],[9E+09,9E+09,9E+09,9E+09,9E+09,9E+09]];
    CONST robtarget Target_4770:=[[-36.104166667,-24.991666667,-2],[0.71519384,0,0,-0.698926156],[0,0,0,0],[9E+09,9E+09,9E+09,9E+09,9E+09,9E+09]];
    CONST robtarget Target_4780:=[[-30.031979167,-28.682604167,-2],[0.71519384,0,0,-0.698926156],[0,0,0,0],[9E+09,9E+09,9E+09,9E+09,9E+09,9E+09]];
    CONST robtarget Target_4790:=[[-25.838333333,-25.785416667,-2],[0.71519384,0,0,-0.698926156],[0,0,0,0],[9E+09,9E+09,9E+09,9E+09,9E+09,9E+09]];
    CONST robtarget Target_4800:=[[-22.875,-25.25625,-2],[0.71519384,0,0,-0.698926156],[0,0,0,0],[9E+09,9E+09,9E+09,9E+09,9E+09,9E+09]];
    CONST robtarget Target_4740:=[[9.563,-21.004,-2],[0.71519384,0,0,-0.698926156],[0,0,0,0],[9E+09,9E+09,9E+09,9E+09,9E+09,9E+09]];
    CONST robtarget Target_4750:=[[6.955,-16.499,-2],[0.71519384,0,0,-0.698926156],[0,0,0,0],[9E+09,9E+09,9E+09,9E+09,9E+09,9E+09]];
    CONST robtarget Target_4730:=[[12.982,-18.059,-2],[0.71519384,0,0,-0.698926156],[0,0,0,0],[9E+09,9E+09,9E+09,9E+09,9E+09,9E+09]];
    CONST robtarget Target_4810:=[[18.929166667,-26.102916667,-2],[0.71519384,0,0,-0.698926156],[0,0,0,0],[9E+09,9E+09,9E+09,9E+09,9E+09,9E+09]];
    CONST robtarget Target_4820:=[[25.093958333,-28.682604167,-2],[0.71519384,0,0,-0.698926156],[0,0,0,0],[9E+09,9E+09,9E+09,9E+09,9E+09,9E+09]];
    CONST robtarget Target_4830:=[[29.089166667,-28.2328125,-2],[0.71519384,0,0,-0.698926156],[0,0,0,0],[9E+09,9E+09,9E+09,9E+09,9E+09,9E+09]];
    CONST robtarget Target_4840:=[[32.455989583,-25.163645833,-2],[0.71519384,0,0,-0.698926156],[0,0,0,0],[9E+09,9E+09,9E+09,9E+09,9E+09,9E+09]];
    CONST robtarget Target_4850:=[[33.745833333,-26.896666667,-2],[0.71519384,0,0,-0.698926156],[0,0,0,0],[9E+09,9E+09,9E+09,9E+09,9E+09,9E+09]];
    CONST robtarget Target_4860:=[[-46.132,-21.991,-2],[0.71519384,0,0,-0.698926156],[0,0,0,0],[9E+09,9E+09,9E+09,9E+09,9E+09,9E+09]];
    CONST robtarget Target_4870:=[[-42.839,-15.759,-2],[0.71519384,0,0,-0.698926156],[0,0,0,0],[9E+09,9E+09,9E+09,9E+09,9E+09,9E+09]];
    CONST robtarget Target_4880:=[[-38.95,-19.202,-2],[0.71519384,0,0,-0.698926156],[0,0,0,0],[9E+09,9E+09,9E+09,9E+09,9E+09,9E+09]];
    CONST robtarget Target_4890:=[[-37.739,-14.66,-2],[0.71519384,0,0,-0.698926156],[0,0,0,0],[9E+09,9E+09,9E+09,9E+09,9E+09,9E+09]];
    CONST robtarget Target_4900:=[[-35.879,-24.873,-2],[0.71519384,0,0,-0.698926156],[0,0,0,0],[9E+09,9E+09,9E+09,9E+09,9E+09,9E+09]];
    CONST robtarget Target_4910:=[[-34.298,-14.146,-2],[0.71519384,0,0,-0.698926156],[0,0,0,0],[9E+09,9E+09,9E+09,9E+09,9E+09,9E+09]];
    CONST robtarget Target_4920:=[[-33.687,-27.261,-2],[0.71519384,0,0,-0.698926156],[0,0,0,0],[9E+09,9E+09,9E+09,9E+09,9E+09,9E+09]];
    CONST robtarget Target_4930:=[[-32.228,-13.941,-2],[0.71519384,0,0,-0.698926156],[0,0,0,0],[9E+09,9E+09,9E+09,9E+09,9E+09,9E+09]];
    CONST robtarget Target_4940:=[[-30.584,-28.667,-2],[0.71519384,0,0,-0.698926156],[0,0,0,0],[9E+09,9E+09,9E+09,9E+09,9E+09,9E+09]];
    CONST robtarget Target_4950:=[[-30.473,-13.878,-2],[0.71519384,0,0,-0.698926156],[0,0,0,0],[9E+09,9E+09,9E+09,9E+09,9E+09,9E+09]];
    CONST robtarget Target_4960:=[[-27.594,-28.036,-2],[0.71519384,0,0,-0.698926156],[0,0,0,0],[9E+09,9E+09,9E+09,9E+09,9E+09,9E+09]];
    CONST robtarget Target_4970:=[[-28.894,-13.755,-2],[0.71519384,0,0,-0.698926156],[0,0,0,0],[9E+09,9E+09,9E+09,9E+09,9E+09,9E+09]];
    CONST robtarget Target_4980:=[[-25.791,-25.62,-2],[0.71519384,0,0,-0.698926156],[0,0,0,0],[9E+09,9E+09,9E+09,9E+09,9E+09,9E+09]];
    CONST robtarget Target_4990:=[[-27.602,-7.296,-2],[0.71519384,0,0,-0.698926156],[0,0,0,0],[9E+09,9E+09,9E+09,9E+09,9E+09,9E+09]];
    CONST robtarget Target_5000:=[[-22.888,-25.241,-2],[0.71519384,0,0,-0.698926156],[0,0,0,0],[9E+09,9E+09,9E+09,9E+09,9E+09,9E+09]];
    CONST robtarget Target_5010:=[[-21.019,-15.317,-2],[0.71519384,0,0,-0.698926156],[0,0,0,0],[9E+09,9E+09,9E+09,9E+09,9E+09,9E+09]];
    CONST robtarget Target_5020:=[[-20.297,-26.307,-2],[0.71519384,0,0,-0.698926156],[0,0,0,0],[9E+09,9E+09,9E+09,9E+09,9E+09,9E+09]];
    CONST robtarget Target_5030:=[[-19.443,-16.447,-2],[0.71519384,0,0,-0.698926156],[0,0,0,0],[9E+09,9E+09,9E+09,9E+09,9E+09,9E+09]];
    CONST robtarget Target_5040:=[[-18.474,-25.262,-2],[0.71519384,0,0,-0.698926156],[0,0,0,0],[9E+09,9E+09,9E+09,9E+09,9E+09,9E+09]];
    CONST robtarget Target_5050:=[[-16.618,-18.319,-2],[0.71519384,0,0,-0.698926156],[0,0,0,0],[9E+09,9E+09,9E+09,9E+09,9E+09,9E+09]];
    CONST robtarget Target_5060:=[[-13.56,-21.394,-2],[0.71519384,0,0,-0.698926156],[0,0,0,0],[9E+09,9E+09,9E+09,9E+09,9E+09,9E+09]];
    CONST robtarget Target_5070:=[[-12.863,-16.193,-2],[0.71519384,0,0,-0.698926156],[0,0,0,0],[9E+09,9E+09,9E+09,9E+09,9E+09,9E+09]];
    CONST robtarget Target_5080:=[[-9.584,-18.831,-2],[0.71519384,0,0,-0.698926156],[0,0,0,0],[9E+09,9E+09,9E+09,9E+09,9E+09,9E+09]];
    CONST robtarget Target_5090:=[[15.754166667,-12.23875,-2],[0.71519384,0,0,-0.698926156],[0,0,0,0],[9E+09,9E+09,9E+09,9E+09,9E+09,9E+09]];
    CONST robtarget Target_5100:=[[12.235208333,-14.71921875,-2],[0.71519384,0,0,-0.698926156],[0,0,0,0],[9E+09,9E+09,9E+09,9E+09,9E+09,9E+09]];
    CONST robtarget Target_5110:=[[7.44625,-16.525,-2],[0.71519384,0,0,-0.698926156],[0,0,0,0],[9E+09,9E+09,9E+09,9E+09,9E+09,9E+09]];
    CONST robtarget Target_5120:=[[5.170833333,-13.82625,-2],[0.71519384,0,0,-0.698926156],[0,0,0,0],[9E+09,9E+09,9E+09,9E+09,9E+09,9E+09]];
    CONST robtarget Target_5130:=[[6.335,-12.609166667,-2],[0.71519384,0,0,-0.698926156],[0,0,0,0],[9E+09,9E+09,9E+09,9E+09,9E+09,9E+09]];
    CONST robtarget Target_5140:=[[-19.329583333,-11.7625,-2],[0.71519384,0,0,-0.698926156],[0,0,0,0],[9E+09,9E+09,9E+09,9E+09,9E+09,9E+09]];
    CONST robtarget Target_5150:=[[-14.031302083,-15.684947917,-2],[0.71519384,0,0,-0.698926156],[0,0,0,0],[9E+09,9E+09,9E+09,9E+09,9E+09,9E+09]];
    CONST robtarget Target_5160:=[[-10.175,-16.789583333,-2],[0.71519384,0,0,-0.698926156],[0,0,0,0],[9E+09,9E+09,9E+09,9E+09,9E+09,9E+09]];
    CONST robtarget Target_5170:=[[-8.534583333,-12.926666667,-2],[0.71519384,0,0,-0.698926156],[0,0,0,0],[9E+09,9E+09,9E+09,9E+09,9E+09,9E+09]];
    ! Posiciones Especiales
    CONST robtarget Target_Home:=[[1.82,196.029178668,-409.843767407],[0.683012702,-0.183012702,-0.183012702,-0.683012702],[0,-1,0,0],[9E+09,9E+09,9E+09,9E+09,9E+09,9E+09]];
    CONST robtarget Target_Pausa:=[[2.8,-2.86,-35.3],[0.71519384,0,0,-0.698926156],[0,0,0,0],[9E+09,9E+09,9E+09,9E+09,9E+09,9E+09]];
    ! Nombres
    CONST robtarget Target_5180:=[[109.688257617,6.242465204,-1.05],[0.71519384,0,0,-0.698926156],[0,0,0,0],[9E+09,9E+09,9E+09,9E+09,9E+09,9E+09]];
    CONST robtarget Target_5190:=[[114.804117077,7.764932412,-1.05],[0.71519384,0,0,-0.698926156],[0,0,0,0],[9E+09,9E+09,9E+09,9E+09,9E+09,9E+09]];
    CONST robtarget Target_5200:=[[114.852149542,14.060921084,-1.05],[0.71519384,0,0,-0.698926156],[0,0,0,0],[9E+09,9E+09,9E+09,9E+09,9E+09,9E+09]];
    CONST robtarget Target_5210:=[[89.788449493,5.806622112,-1.05],[0.71519384,0,0,-0.698926156],[0,0,0,0],[9E+09,9E+09,9E+09,9E+09,9E+09,9E+09]];
    CONST robtarget Target_5220:=[[89.736190172,-1.043413412,-1.05],[0.71519384,0,0,-0.698926156],[0,0,0,0],[9E+09,9E+09,9E+09,9E+09,9E+09,9E+09]];
    CONST robtarget Target_5230:=[[114.671035125,-9.679153857,-1.05],[0.71519384,0,0,-0.698926156],[0,0,0,0],[9E+09,9E+09,9E+09,9E+09,9E+09,9E+09]];
    CONST robtarget Target_5240:=[[114.720348458,-3.21527188,-1.05],[0.71519384,0,0,-0.698926156],[0,0,0,0],[9E+09,9E+09,9E+09,9E+09,9E+09,9E+09]];
    CONST robtarget Target_5250:=[[109.628313096,-1.614929239,-1.05],[0.71519384,0,0,-0.698926156],[0,0,0,0],[9E+09,9E+09,9E+09,9E+09,9E+09,9E+09]];
    CONST robtarget Target_5260:=[[109.688257617,6.242465204,-1.05],[0.71519384,0,0,-0.698926156],[0,0,0,0],[9E+09,9E+09,9E+09,9E+09,9E+09,9E+09]];
    CONST robtarget Target_5270:=[[96.881625508,2.411241866,-1.05],[0.71519384,0,0,-0.698926156],[0,0,0,0],[9E+09,9E+09,9E+09,9E+09,9E+09,9E+09]];
    CONST robtarget Target_5280:=[[105.105704938,-0.20362235,-1.05],[0.71519384,0,0,-0.698926156],[0,0,0,0],[9E+09,9E+09,9E+09,9E+09,9E+09,9E+09]];
    CONST robtarget Target_5290:=[[105.144643255,4.900325652,-1.05],[0.71519384,0,0,-0.698926156],[0,0,0,0],[9E+09,9E+09,9E+09,9E+09,9E+09,9E+09]];
    CONST robtarget Target_5300:=[[96.881625508,2.411241866,-1.05],[0.71519384,0,0,-0.698926156],[0,0,0,0],[9E+09,9E+09,9E+09,9E+09,9E+09,9E+09]];
    CONST robtarget Target_5310:=[[106.487065229,-43.247139436,-1.05],[0.71519384,0,0,-0.698926156],[0,0,0,0],[9E+09,9E+09,9E+09,9E+09,9E+09,9E+09]];
    CONST robtarget Target_5320:=[[98.577300079,-32.240542962,-1.05],[0.71519384,0,0,-0.698926156],[0,0,0,0],[9E+09,9E+09,9E+09,9E+09,9E+09,9E+09]];
    CONST robtarget Target_5330:=[[94.891124892,-34.784882841,-1.05],[0.71519384,0,0,-0.698926156],[0,0,0,0],[9E+09,9E+09,9E+09,9E+09,9E+09,9E+09]];
    CONST robtarget Target_5340:=[[88.328280482,-34.050149,-1.05],[0.71519384,0,0,-0.698926156],[0,0,0,0],[9E+09,9E+09,9E+09,9E+09,9E+09,9E+09]];
    CONST robtarget Target_5350:=[[86.150276379,-31.847995022,-1.05],[0.71519384,0,0,-0.698926156],[0,0,0,0],[9E+09,9E+09,9E+09,9E+09,9E+09,9E+09]];
    CONST robtarget Target_5360:=[[85.266551274,-28.919758171,-1.05],[0.71519384,0,0,-0.698926156],[0,0,0,0],[9E+09,9E+09,9E+09,9E+09,9E+09,9E+09]];
    CONST robtarget Target_5370:=[[86.034650749,-23.822244276,-1.05],[0.71519384,0,0,-0.698926156],[0,0,0,0],[9E+09,9E+09,9E+09,9E+09,9E+09,9E+09]];
    CONST robtarget Target_5380:=[[88.796126234,-14.151711251,-1.05],[0.71519384,0,0,-0.698926156],[0,0,0,0],[9E+09,9E+09,9E+09,9E+09,9E+09,9E+09]];
    CONST robtarget Target_5390:=[[112.835231903,-21.016214048,-1.05],[0.71519384,0,0,-0.698926156],[0,0,0,0],[9E+09,9E+09,9E+09,9E+09,9E+09,9E+09]];
    CONST robtarget Target_5400:=[[111.120258634,-27.021954721,-1.05],[0.71519384,0,0,-0.698926156],[0,0,0,0],[9E+09,9E+09,9E+09,9E+09,9E+09,9E+09]];
    CONST robtarget Target_5410:=[[102.305382668,-24.504816956,-1.05],[0.71519384,0,0,-0.698926156],[0,0,0,0],[9E+09,9E+09,9E+09,9E+09,9E+09,9E+09]];
    CONST robtarget Target_5420:=[[108.589290405,-35.885264197,-1.05],[0.71519384,0,0,-0.698926156],[0,0,0,0],[9E+09,9E+09,9E+09,9E+09,9E+09,9E+09]];
    CONST robtarget Target_5430:=[[106.487065229,-43.247139436,-1.05],[0.71519384,0,0,-0.698926156],[0,0,0,0],[9E+09,9E+09,9E+09,9E+09,9E+09,9E+09]];
    CONST robtarget Target_5440:=[[92.585140666,-28.765895567,-1.05],[0.71519384,0,0,-0.698926156],[0,0,0,0],[9E+09,9E+09,9E+09,9E+09,9E+09,9E+09]];
    CONST robtarget Target_5450:=[[96.721165901,-27.092100996,-1.05],[0.71519384,0,0,-0.698926156],[0,0,0,0],[9E+09,9E+09,9E+09,9E+09,9E+09,9E+09]];
    CONST robtarget Target_5460:=[[97.978666438,-23.269298627,-1.05],[0.71519384,0,0,-0.698926156],[0,0,0,0],[9E+09,9E+09,9E+09,9E+09,9E+09,9E+09]];
    CONST robtarget Target_5470:=[[91.504736215,-21.42063118,-1.05],[0.71519384,0,0,-0.698926156],[0,0,0,0],[9E+09,9E+09,9E+09,9E+09,9E+09,9E+09]];
    CONST robtarget Target_5480:=[[90.446913725,-26.531447268,-1.05],[0.71519384,0,0,-0.698926156],[0,0,0,0],[9E+09,9E+09,9E+09,9E+09,9E+09,9E+09]];
    CONST robtarget Target_5490:=[[91.126319123,-27.973910396,-1.05],[0.71519384,0,0,-0.698926156],[0,0,0,0],[9E+09,9E+09,9E+09,9E+09,9E+09,9E+09]];
    CONST robtarget Target_5500:=[[93.095027208,-58.892961182,-1.05],[0.714513134,0.030486731,0.031196317,-0.698260933],[0,0,0,0],[9E+09,9E+09,9E+09,9E+09,9E+09,9E+09]];
    CONST robtarget Target_5510:=[[78.975116655,-50.810976236,-1.05],[0.714513134,0.030486731,0.031196317,-0.698260933],[0,0,0,0],[9E+09,9E+09,9E+09,9E+09,9E+09,9E+09]];
    CONST robtarget Target_5520:=[[77.190240488,-53.929305705,-1.05],[0.714513134,0.030486731,0.031196317,-0.698260933],[0,0,0,0],[9E+09,9E+09,9E+09,9E+09,9E+09,9E+09]];
    CONST robtarget Target_5530:=[[73.401615648,-51.760764424,-1.05],[0.714513134,0.030486731,0.031196317,-0.698260933],[0,0,0,0],[9E+09,9E+09,9E+09,9E+09,9E+09,9E+09]];
    CONST robtarget Target_5540:=[[80.090730499,-40.07431561,-1.05],[0.714513134,0.030486731,0.031196317,-0.698260933],[0,0,0,0],[9E+09,9E+09,9E+09,9E+09,9E+09,9E+09]];
    CONST robtarget Target_5550:=[[83.87935534,-42.242856892,-1.05],[0.714513134,0.030486731,0.031196317,-0.698260933],[0,0,0,0],[9E+09,9E+09,9E+09,9E+09,9E+09,9E+09]];
    CONST robtarget Target_5560:=[[82.094479173,-45.361186361,-1.05],[0.714513134,0.030486731,0.031196317,-0.698260933],[0,0,0,0],[9E+09,9E+09,9E+09,9E+09,9E+09,9E+09]];
    CONST robtarget Target_5570:=[[96.214389726,-53.443171307,-1.05],[0.714513134,0.030486731,0.031196317,-0.698260933],[0,0,0,0],[9E+09,9E+09,9E+09,9E+09,9E+09,9E+09]];
    CONST robtarget Target_5580:=[[97.999265893,-50.324841838,-1.05],[0.714513134,0.030486731,0.031196317,-0.698260933],[0,0,0,0],[9E+09,9E+09,9E+09,9E+09,9E+09,9E+09]];
    CONST robtarget Target_5590:=[[101.787890733,-52.49338312,-1.05],[0.714513134,0.030486731,0.031196317,-0.698260933],[0,0,0,0],[9E+09,9E+09,9E+09,9E+09,9E+09,9E+09]];
    CONST robtarget Target_5600:=[[95.098775882,-64.179831933,-1.05],[0.714513134,0.030486731,0.031196317,-0.698260933],[0,0,0,0],[9E+09,9E+09,9E+09,9E+09,9E+09,9E+09]];
    CONST robtarget Target_5610:=[[91.310151041,-62.011290651,-1.05],[0.714513134,0.030486731,0.031196317,-0.698260933],[0,0,0,0],[9E+09,9E+09,9E+09,9E+09,9E+09,9E+09]];
    CONST robtarget Target_5620:=[[93.095027208,-58.892961182,-1.05],[0.714513134,0.030486731,0.031196317,-0.698260933],[0,0,0,0],[9E+09,9E+09,9E+09,9E+09,9E+09,9E+09]];
    CONST robtarget Target_5630:=[[87.599014409,-74.670979869,-1.05],[0.709075258,0.09122817,0.093351528,-0.692946745],[0,0,0,0],[9E+09,9E+09,9E+09,9E+09,9E+09,9E+09]];
    CONST robtarget Target_5640:=[[69.19067617,-57.755511112,-1.05],[0.709075258,0.09122817,0.093351528,-0.692946745],[0,0,0,0],[9E+09,9E+09,9E+09,9E+09,9E+09,9E+09]];
    CONST robtarget Target_5650:=[[57.750866224,-70.204937959,-1.05],[0.709075258,0.09122817,0.093351528,-0.692946745],[0,0,0,0],[9E+09,9E+09,9E+09,9E+09,9E+09,9E+09]];
    CONST robtarget Target_5660:=[[61.26192719,-73.431260797,-1.05],[0.709075258,0.09122817,0.093351528,-0.692946745],[0,0,0,0],[9E+09,9E+09,9E+09,9E+09,9E+09,9E+09]];
    CONST robtarget Target_5670:=[[68.475709757,-65.580828073,-1.05],[0.709075258,0.09122817,0.093351528,-0.692946745],[0,0,0,0],[9E+09,9E+09,9E+09,9E+09,9E+09,9E+09]];
    CONST robtarget Target_5680:=[[71.70242245,-68.545862561,-1.05],[0.709075258,0.09122817,0.093351528,-0.692946745],[0,0,0,0],[9E+09,9E+09,9E+09,9E+09,9E+09,9E+09]];
    CONST robtarget Target_5690:=[[65.056654353,-75.778150873,-1.05],[0.709075258,0.09122817,0.093351528,-0.692946745],[0,0,0,0],[9E+09,9E+09,9E+09,9E+09,9E+09,9E+09]];
    CONST robtarget Target_5700:=[[68.567712686,-79.004471291,-1.05],[0.709075258,0.09122817,0.093351528,-0.692946745],[0,0,0,0],[9E+09,9E+09,9E+09,9E+09,9E+09,9E+09]];
    CONST robtarget Target_5710:=[[75.213480783,-71.77218298,-1.05],[0.709075258,0.09122817,0.093351528,-0.692946745],[0,0,0,0],[9E+09,9E+09,9E+09,9E+09,9E+09,9E+09]];
    CONST robtarget Target_5720:=[[79.861927819,-76.043652767,-1.05],[0.709075258,0.09122817,0.093351528,-0.692946745],[0,0,0,0],[9E+09,9E+09,9E+09,9E+09,9E+09,9E+09]];
    CONST robtarget Target_5730:=[[72.648145252,-83.894085491,-1.05],[0.709075258,0.09122817,0.093351528,-0.692946745],[0,0,0,0],[9E+09,9E+09,9E+09,9E+09,9E+09,9E+09]];
    CONST robtarget Target_5740:=[[76.159204462,-87.120406716,-1.05],[0.709075258,0.09122817,0.093351528,-0.692946745],[0,0,0,0],[9E+09,9E+09,9E+09,9E+09,9E+09,9E+09]];
    CONST robtarget Target_5750:=[[87.599014409,-74.670979869,-1.05],[0.709075258,0.09122817,0.093351528,-0.692946745],[0,0,0,0],[9E+09,9E+09,9E+09,9E+09,9E+09,9E+09]];
    CONST robtarget Target_5760:=[[52.229331861,-74.691344254,-1.05],[0.709075258,0.09122817,0.093351528,-0.692946745],[0,0,0,0],[9E+09,9E+09,9E+09,9E+09,9E+09,9E+09]];
    CONST robtarget Target_5770:=[[47.018436392,-78.195228433,-1.05],[0.709075258,0.09122817,0.093351528,-0.692946745],[0,0,0,0],[9E+09,9E+09,9E+09,9E+09,9E+09,9E+09]];
    CONST robtarget Target_5780:=[[58.307689931,-94.98434506,-1.05],[0.709075258,0.09122817,0.093351528,-0.692946745],[0,0,0,0],[9E+09,9E+09,9E+09,9E+09,9E+09,9E+09]];
    CONST robtarget Target_5790:=[[49.669306498,-100.792923493,-1.05],[0.709075258,0.09122817,0.093351528,-0.692946745],[0,0,0,0],[9E+09,9E+09,9E+09,9E+09,9E+09,9E+09]];
    CONST robtarget Target_5800:=[[52.330009674,-104.749859686,-1.05],[0.709075258,0.09122817,0.093351528,-0.692946745],[0,0,0,0],[9E+09,9E+09,9E+09,9E+09,9E+09,9E+09]];
    CONST robtarget Target_5810:=[[66.179288577,-95.437397075,-1.05],[0.709075258,0.09122817,0.093351528,-0.692946745],[0,0,0,0],[9E+09,9E+09,9E+09,9E+09,9E+09,9E+09]];
    CONST robtarget Target_5820:=[[52.229331861,-74.691344254,-1.05],[0.709075258,0.09122817,0.093351528,-0.692946745],[0,0,0,0],[9E+09,9E+09,9E+09,9E+09,9E+09,9E+09]];
    CONST robtarget Target_5830:=[[-55.053122352,-94.880976532,-1.05],[0.709075257,0.09122817,0.093351529,-0.692946746],[0,0,0,0],[9E+09,9E+09,9E+09,9E+09,9E+09,9E+09]];
    CONST robtarget Target_5840:=[[-57.04231561,-97.259064884,-1.05],[0.709075257,0.09122817,0.093351529,-0.692946746],[0,0,0,0],[9E+09,9E+09,9E+09,9E+09,9E+09,9E+09]];
    CONST robtarget Target_5850:=[[-61.029786691,-96.378761325,-1.05],[0.709075257,0.09122817,0.093351529,-0.692946746],[0,0,0,0],[9E+09,9E+09,9E+09,9E+09,9E+09,9E+09]];
    CONST robtarget Target_5860:=[[-52.627930216,-77.202859768,-1.05],[0.709075257,0.09122817,0.093351529,-0.692946746],[0,0,0,0],[9E+09,9E+09,9E+09,9E+09,9E+09,9E+09]];
    CONST robtarget Target_5870:=[[-57.062793404,-74.828016046,-1.05],[0.709075257,0.09122817,0.093351529,-0.692946746],[0,0,0,0],[9E+09,9E+09,9E+09,9E+09,9E+09,9E+09]];
    CONST robtarget Target_5880:=[[-65.709323186,-91.263830896,-1.05],[0.709075257,0.09122817,0.093351529,-0.692946746],[0,0,0,0],[9E+09,9E+09,9E+09,9E+09,9E+09,9E+09]];
    CONST robtarget Target_5890:=[[-66.325791382,-95.467544737,-1.05],[0.709075257,0.09122817,0.093351529,-0.692946746],[0,0,0,0],[9E+09,9E+09,9E+09,9E+09,9E+09,9E+09]];
    CONST robtarget Target_5900:=[[-64.114177839,-99.519648554,-1.05],[0.709075257,0.09122817,0.093351529,-0.692946746],[0,0,0,0],[9E+09,9E+09,9E+09,9E+09,9E+09,9E+09]];
    CONST robtarget Target_5910:=[[-58.628621279,-102.244344742,-1.05],[0.709075257,0.09122817,0.093351529,-0.692946746],[0,0,0,0],[9E+09,9E+09,9E+09,9E+09,9E+09,9E+09]];
    CONST robtarget Target_5920:=[[-53.230803989,-100.472859457,-1.05],[0.709075257,0.09122817,0.093351529,-0.692946746],[0,0,0,0],[9E+09,9E+09,9E+09,9E+09,9E+09,9E+09]];
    CONST robtarget Target_5930:=[[-51.116403585,-97.608084827,-1.05],[0.709075257,0.09122817,0.093351529,-0.692946746],[0,0,0,0],[9E+09,9E+09,9E+09,9E+09,9E+09,9E+09]];
    CONST robtarget Target_5940:=[[-55.053122352,-94.880976532,-1.05],[0.709075257,0.09122817,0.093351529,-0.692946746],[0,0,0,0],[9E+09,9E+09,9E+09,9E+09,9E+09,9E+09]];
    CONST robtarget Target_5950:=[[-67.578159329,-66.268206974,-1.05],[0.709075257,0.09122817,0.093351529,-0.692946746],[0,0,0,0],[9E+09,9E+09,9E+09,9E+09,9E+09,9E+09]];
    CONST robtarget Target_5960:=[[-78.425488647,-90.806992983,-1.05],[0.709075257,0.09122817,0.093351529,-0.692946746],[0,0,0,0],[9E+09,9E+09,9E+09,9E+09,9E+09,9E+09]];
    CONST robtarget Target_5970:=[[-82.203341971,-87.012166569,-1.05],[0.709075257,0.09122817,0.093351529,-0.692946746],[0,0,0,0],[9E+09,9E+09,9E+09,9E+09,9E+09,9E+09]];
    CONST robtarget Target_5980:=[[-79.634688759,-81.54337923,-1.05],[0.709075257,0.09122817,0.093351529,-0.692946746],[0,0,0,0],[9E+09,9E+09,9E+09,9E+09,9E+09,9E+09]];
    CONST robtarget Target_5990:=[[-86.685077169,-74.461314929,-1.05],[0.709075257,0.09122817,0.093351529,-0.692946746],[0,0,0,0],[9E+09,9E+09,9E+09,9E+09,9E+09,9E+09]];
    CONST robtarget Target_6000:=[[-92.249543825,-76.920829274,-1.05],[0.709075257,0.09122817,0.093351529,-0.692946746],[0,0,0,0],[9E+09,9E+09,9E+09,9E+09,9E+09,9E+09]];
    CONST robtarget Target_6010:=[[-96.123648503,-73.02931907,-1.05],[0.709075257,0.09122817,0.093351529,-0.692946746],[0,0,0,0],[9E+09,9E+09,9E+09,9E+09,9E+09,9E+09]];
    CONST robtarget Target_6020:=[[-71.343981497,-62.48546577,-1.05],[0.709075257,0.09122817,0.093351529,-0.692946746],[0,0,0,0],[9E+09,9E+09,9E+09,9E+09,9E+09,9E+09]];
    CONST robtarget Target_6030:=[[-67.578159329,-66.268206974,-1.05],[0.709075257,0.09122817,0.093351529,-0.692946746],[0,0,0,0],[9E+09,9E+09,9E+09,9E+09,9E+09,9E+09]];
    CONST robtarget Target_6040:=[[-82.556994559,-72.637680689,-1.05],[0.709075257,0.09122817,0.093351529,-0.692946746],[0,0,0,0],[9E+09,9E+09,9E+09,9E+09,9E+09,9E+09]];
    CONST robtarget Target_6050:=[[-73.552178938,-68.533867673,-1.05],[0.709075257,0.09122817,0.093351529,-0.692946746],[0,0,0,0],[9E+09,9E+09,9E+09,9E+09,9E+09,9E+09]];
    CONST robtarget Target_6060:=[[-77.744442443,-77.471854575,-1.05],[0.709075257,0.09122817,0.093351529,-0.692946746],[0,0,0,0],[9E+09,9E+09,9E+09,9E+09,9E+09,9E+09]];
    CONST robtarget Target_6070:=[[-82.556994559,-72.637680689,-1.05],[0.709075257,0.09122817,0.093351529,-0.692946746],[0,0,0,0],[9E+09,9E+09,9E+09,9E+09,9E+09,9E+09]];
    CONST robtarget Target_6080:=[[-102.323579234,-63.695242302,-1.05],[0.709075257,0.09122817,0.093351529,-0.692946746],[0,0,0,0],[9E+09,9E+09,9E+09,9E+09,9E+09,9E+09]];
    CONST robtarget Target_6090:=[[-79.913220601,-52.614816952,-1.05],[0.709075257,0.09122817,0.093351529,-0.692946746],[0,0,0,0],[9E+09,9E+09,9E+09,9E+09,9E+09,9E+09]];
    CONST robtarget Target_6100:=[[-86.306364197,-40.064519811,-1.05],[0.709075257,0.09122817,0.093351529,-0.692946746],[0,0,0,0],[9E+09,9E+09,9E+09,9E+09,9E+09,9E+09]];
    CONST robtarget Target_6110:=[[-89.370507714,-37.118454493,-1.05],[0.709075257,0.09122817,0.093351529,-0.692946746],[0,0,0,0],[9E+09,9E+09,9E+09,9E+09,9E+09,9E+09]];
    CONST robtarget Target_6120:=[[-93.261057975,-36.70927707,-1.05],[0.709075257,0.09122817,0.093351529,-0.692946746],[0,0,0,0],[9E+09,9E+09,9E+09,9E+09,9E+09,9E+09]];
    CONST robtarget Target_6130:=[[-97.377714772,-38.901635279,-1.05],[0.709075257,0.09122817,0.093351529,-0.692946746],[0,0,0,0],[9E+09,9E+09,9E+09,9E+09,9E+09,9E+09]];
    CONST robtarget Target_6140:=[[-99.115871381,-43.446898875,-1.05],[0.709075257,0.09122817,0.093351529,-0.692946746],[0,0,0,0],[9E+09,9E+09,9E+09,9E+09,9E+09,9E+09]];
    CONST robtarget Target_6150:=[[-112.285380271,-43.54732137,-1.05],[0.709075257,0.09122817,0.093351529,-0.692946746],[0,0,0,0],[9E+09,9E+09,9E+09,9E+09,9E+09,9E+09]];
    CONST robtarget Target_6160:=[[-109.609752413,-48.958826611,-1.05],[0.709075257,0.09122817,0.093351529,-0.692946746],[0,0,0,0],[9E+09,9E+09,9E+09,9E+09,9E+09,9E+09]];
    CONST robtarget Target_6170:=[[-98.64243137,-50.575023886,-1.05],[0.709075257,0.09122817,0.093351529,-0.692946746],[0,0,0,0],[9E+09,9E+09,9E+09,9E+09,9E+09,9E+09]];
    CONST robtarget Target_6180:=[[-95.205344109,-54.544706786,-1.05],[0.709075257,0.09122817,0.093351529,-0.692946746],[0,0,0,0],[9E+09,9E+09,9E+09,9E+09,9E+09,9E+09]];
    CONST robtarget Target_6190:=[[-104.560827202,-59.170368237,-1.05],[0.709075257,0.09122817,0.093351529,-0.692946746],[0,0,0,0],[9E+09,9E+09,9E+09,9E+09,9E+09,9E+09]];
    CONST robtarget Target_6200:=[[-102.323579234,-63.695242302,-1.05],[0.709075257,0.09122817,0.093351529,-0.692946746],[0,0,0,0],[9E+09,9E+09,9E+09,9E+09,9E+09,9E+09]];
    CONST robtarget Target_6210:=[[-85.941579742,-49.964394118,-1.05],[0.709075257,0.09122817,0.093351529,-0.692946746],[0,0,0,0],[9E+09,9E+09,9E+09,9E+09,9E+09,9E+09]];
    CONST robtarget Target_6220:=[[-89.396560283,-43.169013101,-1.05],[0.709075257,0.09122817,0.093351529,-0.692946746],[0,0,0,0],[9E+09,9E+09,9E+09,9E+09,9E+09,9E+09]];
    CONST robtarget Target_6230:=[[-93.243612809,-42.198530228,-1.05],[0.709075257,0.09122817,0.093351529,-0.692946746],[0,0,0,0],[9E+09,9E+09,9E+09,9E+09,9E+09,9E+09]];
    CONST robtarget Target_6240:=[[-95.018846426,-45.225953832,-1.05],[0.709075257,0.09122817,0.093351529,-0.692946746],[0,0,0,0],[9E+09,9E+09,9E+09,9E+09,9E+09,9E+09]];
    CONST robtarget Target_6250:=[[-91.628246501,-52.776070966,-1.05],[0.709075257,0.09122817,0.093351529,-0.692946746],[0,0,0,0],[9E+09,9E+09,9E+09,9E+09,9E+09,9E+09]];
    CONST robtarget Target_6260:=[[-85.941579742,-49.964394118,-1.05],[0.709075257,0.09122817,0.093351529,-0.692946746],[0,0,0,0],[9E+09,9E+09,9E+09,9E+09,9E+09,9E+09]];
    CONST robtarget Target_6270:=[[-115.123528363,-32.683782748,-1.05],[0.71519384,0,0,-0.698926156],[0,0,0,0],[9E+09,9E+09,9E+09,9E+09,9E+09,9E+09]];
    CONST robtarget Target_6280:=[[-90.384106581,-29.083642487,-1.05],[0.71519384,0,0,-0.698926156],[0,0,0,0],[9E+09,9E+09,9E+09,9E+09,9E+09,9E+09]];
    CONST robtarget Target_6290:=[[-93.053514695,-10.740020174,-1.05],[0.71519384,0,0,-0.698926156],[0,0,0,0],[9E+09,9E+09,9E+09,9E+09,9E+09,9E+09]];
    CONST robtarget Target_6300:=[[-97.238628367,-11.349047999,-1.05],[0.71519384,0,0,-0.698926156],[0,0,0,0],[9E+09,9E+09,9E+09,9E+09,9E+09,9E+09]];
    CONST robtarget Target_6310:=[[-95.296124385,-24.697534961,-1.05],[0.71519384,0,0,-0.698926156],[0,0,0,0],[9E+09,9E+09,9E+09,9E+09,9E+09,9E+09]];
    CONST robtarget Target_6320:=[[-100.78064895,-25.495656189,-1.05],[0.71519384,0,0,-0.698926156],[0,0,0,0],[9E+09,9E+09,9E+09,9E+09,9E+09,9E+09]];
    CONST robtarget Target_6330:=[[-102.588086216,-13.075319865,-1.05],[0.71519384,0,0,-0.698926156],[0,0,0,0],[9E+09,9E+09,9E+09,9E+09,9E+09,9E+09]];
    CONST robtarget Target_6340:=[[-106.756323565,-13.681891807,-1.05],[0.71519384,0,0,-0.698926156],[0,0,0,0],[9E+09,9E+09,9E+09,9E+09,9E+09,9E+09]];
    CONST robtarget Target_6350:=[[-104.948886299,-26.102228131,-1.05],[0.71519384,0,0,-0.698926156],[0,0,0,0],[9E+09,9E+09,9E+09,9E+09,9E+09,9E+09]];
    CONST robtarget Target_6360:=[[-111.682195145,-27.082075456,-1.05],[0.71519384,0,0,-0.698926156],[0,0,0,0],[9E+09,9E+09,9E+09,9E+09,9E+09,9E+09]];
    CONST robtarget Target_6370:=[[-113.693460428,-13.261075014,-1.05],[0.71519384,0,0,-0.698926156],[0,0,0,0],[9E+09,9E+09,9E+09,9E+09,9E+09,9E+09]];
    CONST robtarget Target_6380:=[[-117.861697776,-13.867646955,-1.05],[0.71519384,0,0,-0.698926156],[0,0,0,0],[9E+09,9E+09,9E+09,9E+09,9E+09,9E+09]];
    CONST robtarget Target_6390:=[[-115.123528363,-32.683782748,-1.05],[0.71519384,0,0,-0.698926156],[0,0,0,0],[9E+09,9E+09,9E+09,9E+09,9E+09,9E+09]];
    CONST robtarget Target_6400:=[[-117.726404557,-1.136381061,-1.05],[0.71519384,0,0,-0.698926156],[0,0,0,0],[9E+09,9E+09,9E+09,9E+09,9E+09,9E+09]];
    CONST robtarget Target_6410:=[[-93.087497101,-5.370083856,-1.05],[0.71519384,0,0,-0.698926156],[0,0,0,0],[9E+09,9E+09,9E+09,9E+09,9E+09,9E+09]];
    CONST robtarget Target_6420:=[[-91.177098035,6.45277272,-1.05],[0.71519384,0,0,-0.698926156],[0,0,0,0],[9E+09,9E+09,9E+09,9E+09,9E+09,9E+09]];
    CONST robtarget Target_6430:=[[-91.730723643,10.65739529,-1.05],[0.71519384,0,0,-0.698926156],[0,0,0,0],[9E+09,9E+09,9E+09,9E+09,9E+09,9E+09]];
    CONST robtarget Target_6440:=[[-94.399809505,14.269519799,-1.05],[0.71519384,0,0,-0.698926156],[0,0,0,0],[9E+09,9E+09,9E+09,9E+09,9E+09,9E+09]];
    CONST robtarget Target_6450:=[[-102.092983713,17.442872972,-1.05],[0.71519384,0,0,-0.698926156],[0,0,0,0],[9E+09,9E+09,9E+09,9E+09,9E+09,9E+09]];
    CONST robtarget Target_6460:=[[-107.466692974,17.587595318,-1.05],[0.71519384,0,0,-0.698926156],[0,0,0,0],[9E+09,9E+09,9E+09,9E+09,9E+09,9E+09]];
    CONST robtarget Target_6470:=[[-112.273081014,15.696886799,-1.05],[0.71519384,0,0,-0.698926156],[0,0,0,0],[9E+09,9E+09,9E+09,9E+09,9E+09,9E+09]];
    CONST robtarget Target_6480:=[[-114.84017674,12.538939522,-1.05],[0.71519384,0,0,-0.698926156],[0,0,0,0],[9E+09,9E+09,9E+09,9E+09,9E+09,9E+09]];
    CONST robtarget Target_6490:=[[-116.117828616,8.225058717,-1.05],[0.71519384,0,0,-0.698926156],[0,0,0,0],[9E+09,9E+09,9E+09,9E+09,9E+09,9E+09]];
    CONST robtarget Target_6500:=[[-117.726404557,-1.136381061,-1.05],[0.71519384,0,0,-0.698926156],[0,0,0,0],[9E+09,9E+09,9E+09,9E+09,9E+09,9E+09]];
    CONST robtarget Target_6510:=[[-112.72027567,3.12514161,-1.05],[0.71519384,0,0,-0.698926156],[0,0,0,0],[9E+09,9E+09,9E+09,9E+09,9E+09,9E+09]];
    CONST robtarget Target_6520:=[[-96.400780227,0.320963153,-1.05],[0.71519384,0,0,-0.698926156],[0,0,0,0],[9E+09,9E+09,9E+09,9E+09,9E+09,9E+09]];
    CONST robtarget Target_6530:=[[-95.550216265,6.68078536,-1.05],[0.71519384,0,0,-0.698926156],[0,0,0,0],[9E+09,9E+09,9E+09,9E+09,9E+09,9E+09]];
    CONST robtarget Target_6540:=[[-98.458238684,11.004462137,-1.05],[0.71519384,0,0,-0.698926156],[0,0,0,0],[9E+09,9E+09,9E+09,9E+09,9E+09,9E+09]];
    CONST robtarget Target_6550:=[[-102.758200984,12.262418381,-1.05],[0.71519384,0,0,-0.698926156],[0,0,0,0],[9E+09,9E+09,9E+09,9E+09,9E+09,9E+09]];
    CONST robtarget Target_6560:=[[-107.357490113,12.533620267,-1.05],[0.71519384,0,0,-0.698926156],[0,0,0,0],[9E+09,9E+09,9E+09,9E+09,9E+09,9E+09]];
    CONST robtarget Target_6570:=[[-111.32980761,9.807467907,-1.05],[0.71519384,0,0,-0.698926156],[0,0,0,0],[9E+09,9E+09,9E+09,9E+09,9E+09,9E+09]];
    CONST robtarget Target_6580:=[[-112.72027567,3.12514161,-1.05],[0.71519384,0,0,-0.698926156],[0,0,0,0],[9E+09,9E+09,9E+09,9E+09,9E+09,9E+09]];

    !Tiempos de la banda
    CONST num TiempoEntrada := 4.3;
    CONST num TiempoSalida := 4.3;

    ! Pose de mantenimiento y de farmeo de aura
    CONST jointtarget PoseMant :=[[-30,-10,10,0,30,0],[9E+09,9E+09,9E+09,9E+09,9E+09,9E+09]];
    CONST robtarget Pivote:=[[-2.796,3.031,-102],[0.707106781,0,0,-0.707106781],[0,0,0,0],[9E+09,9E+09,9E+09,9E+09,9E+09,9E+09]];
    CONST jointtarget Pose_Aura1:=[[-9.97,22.69,-26.9,14.96,-6,-2.72],[9E+09,9E+09,9E+09,9E+09,9E+09,9E+09]];
    CONST jointtarget Pose_Aura2:=[[10,15,-10,0,20,0],[9E+09,9E+09,9E+09,9E+09,9E+09,9E+09]];
    CONST jointtarget Pose_Aura3:=[[10,25,-5,0,30,0],[9E+09,9E+09,9E+09,9E+09,9E+09,9E+09]];
    CONST jointtarget Pose_Aura4:=[[-20.82,-13.81,1.11,0,5.28,95.41],[9E+09,9E+09,9E+09,9E+09,9E+09,9E+09]];
    CONST num TiempoDeslizamiento:=3.8;




    PROC main()
        Reset DO_01;
        Reset DO_02;
        Reset DO_03;
        ConveyorStop;
        Path_Home;

        WHILE TRUE DO

            IF DI_01=1 THEN
                CicloDecoracion;
            ENDIF

            IF DI_02 = 1 THEN
                ConveyorStop;
                Set DO_02;
                Path_Home;
                WHILE DI_02 = 0 DO
                    ModoMantenimiento;
                ENDWHILE
                Path_Home;
                Reset DO_02;
            ENDIF

            IF DI_03 = 1 THEN
                ConveyorStop;
                Set DO_03;
                FarmearAura;
                Reset DO_03;
            ENDIF

        ENDWHILE
    ENDPROC




    PROC RutinaVuelta()
        IF DI_02 = 1 THEN
            Path_Home;
            ConveyorBackward;
            WaitTime 4.3;
            ConveyorStop;
        ENDIF
    ENDPROC


PROC RutinaDecoracion()

        ! Contornos principales y rostro
        Path_Home;
        Path_ContornoExterno; !1
        Path_Pausa;
        Path_Cabello; !2
        Path_Pausa;
        Path_ContornoCara; !3
        Path_Pausa;
        Path_Frente; !4
        Path_Pausa;
        Path_Boca; !5
        Path_Pausa;

        ! Elementos Ninja
        Path_BandaNinja; !6
        Path_Pausa;
        Path_SimboloNinja; !7
        Path_Pausa;

        ! Orejas
        Path_OrejaDerecha1; !8
        Path_Pausa;
        Path_OrejaDerecha2; !9
        Path_Pausa;
        Path_OrejaIzquierda1; !10
        Path_Pausa;
        Path_OrejaIzquierda2; !11
        Path_Pausa;

        ! Detalles
        Path_Detalle1; !12
        Path_Pausa;
        Path_Detalle2; !13
        Path_Pausa;
        Path_Detalle3; !14
        Path_Pausa;
        Path_Detalle4; !15
        Path_Pausa;
        Path_Detalle5; !16
        Path_Pausa;
        Path_Detalle6; !17
        Path_Pausa;
        Path_Detalle7; !18
        Path_Pausa;

        ! Nombre 1: ARIEL
        Path_Nombre1_A1; !19
        Path_Pausa;
        Path_Nombre1_A2; !20
        Path_Pausa;
        Path_Nombre1_R1; !21
        Path_Pausa;
        Path_Nombre1_R2; !22
        Path_Pausa;
        Path_Nombre1_I; !23
        Path_Pausa;
        Path_Nombre1_E; !24
        Path_Pausa;
        Path_Nombre1_L; !25
        Path_Pausa;

        ! Nombre 2: JARED
        Path_Nombre2_J; !26
        Path_Pausa;
        Path_Nombre2_A1; !27
        Path_Pausa;
        Path_Nombre2_A2; !28
        Path_Pausa;
        Path_Nombre2_R1; !29
        Path_Pausa;
        Path_Nombre2_R2; !30
        Path_Pausa;
        Path_Nombre2_E; !31
        Path_Pausa;
        Path_Nombre2_D1; !32
        Path_Pausa;
        Path_Nombre2_D2; !33
        Path_Pausa;

        ! Pintado final
        Path_Pintar1; !34
        Path_Pausa;
        Path_Pintar2; !35
        Path_Pausa;
        Path_Home;

ENDPROC

PROC ModoMantenimiento()
    MoveAbsJ PoseMant, v200, fine, MyNewTool;
ENDPROC

PROC FarmearAura()
    VAR num i;
    Reset DO_01;
    Reset DO_02;
    Set DO_03;

    Path_Home;


    MoveAbsJ Pose_Aura1, v150, z1, MyNewTool;

    FOR i FROM 1 TO 3 DO
        MoveAbsJ Pose_Aura2, v150, z1, MyNewTool;
        MoveAbsJ Pose_Aura3, v150, z1, MyNewTool;
    ENDFOR

    MoveAbsJ Pose_Aura4, v150, fine, MyNewTool;
    Path_Home;
    Reset DO_03;

    WHILE DI_03 = 1 DO
        WaitTime 0.1;
    ENDWHILE
ENDPROC

